  rq_init_comm_if_connected(9, "1")
  rq_init_comm_if_connected(2, "2")
  rq_init_comm_if_connected(3, "3")
  rq_init_comm_if_connected(4, "4")
  rq_print_connected_grippers()
  rq_gripper_communication_thread = run rq_gripper_communication()
  set_closed_norm(97.6470588235294, 1)
  set_open_norm(1.1764705882352942, 1)
  set_closed_mm(0.0, 1)
  set_open_mm(53.0, 1)
  set_closed_norm(100.0, 2)
  set_open_norm(0.0, 2)
  set_closed_mm(0.0, 2)
  set_open_mm(50.0, 2)
  set_closed_norm(100.0, 3)
  set_open_norm(0.0, 3)
  set_closed_mm(0.0, 3)
  set_open_mm(50.0, 3)
  set_closed_norm(100.0, 4)
  set_open_norm(0.0, 4)
  set_closed_mm(0.0, 4)
  set_open_mm(50.0, 4)
  rq_current_limit_enabled = False
  while(not rq_gripper_communication_thread_started):
      sync()
  end
  # end: URCap Installation Node
  global AMR_Position=struct(position_identifier=0, x1=0, x2=0, y1=0, y2=0, theta1=0, theta2=0)
  global CAM_Pose=p[0,0,0,0,0,0]
  global CAM_Relation=""
  global CMD_Abort=  False
  global CMD_Clear=  False
  global CMD_Reset=  False
  global CMD_Start=  False
  global CMD_Suspend=  False
  global CMD_Unhold=  False
  global CMD_Unsuspend=  False
  global CNT_Rack_Output=0
  global FNC_Freedrive=  False
  global PRC_TubCounter=0
  global PRC_TubNumber=0
  global STP=0
  global TMR_Barcode=0
  global TMR_Barcode_is_counting=False
  thread Timer_Thread():
    while (True):
      if (TMR_Barcode_is_counting):
        TMR_Barcode = TMR_Barcode + get_steptime()
      end
      sync()
    end
  end
  run Timer_Thread()
  def Sub_Vision_V18():
    $ 698 "Sub_Vision_V18" "noBreak"
    $ 699 "PreSettings"
    $ 700 "CAM_LM_Detected≔ False "
    global CAM_LM_Detected=  False
    $ 701 "CAM_Captures≔0"
    global CAM_Captures=0
    $ 702 "CAM_Pose≔p[0,0,0,0,0,0]"
    global CAM_Pose=p[0,0,0,0,0,0]
    $ 703 "CAM_LM_Refinmnt≔ False "
    global CAM_LM_Refinmnt=  False
    $ 704 "CAM_LM_Refined≔ False "
    global CAM_LM_Refined=  False
    $ 705 "CAM_LM_Deviatn≔p[0,0,0,0,0,0]"
    global CAM_LM_Deviatn=p[0,0,0,0,0,0]
    $ 706 "CAM_LM_ID≔0"
    global CAM_LM_ID=0
    $ 707 "CAM_Done≔ False "
    global CAM_Done=  False
    $ 708 "CAM_CNT_Obj≔0"
    global CAM_CNT_Obj=0
    $ 709 "CAM_Result = []"
    CAM_Result = []
    $ 710 "OBJ_Detected≔ False "
    global OBJ_Detected=  False
    $ 711 "FRM_Reference≔p[0,0,0,0,0,0]"
    global FRM_Reference=p[0,0,0,0,0,0]
    $ 712 "'=========='"
    # '=========='
    $ 713 "Switch Action"
    switch_1 = Action
    $ 714 "Case 13"
    if (13 == switch_1):
    elif (15 == switch_1):
      $ 832 "Case 15"
    elif (131 == switch_1):
      $ 878 "Case 131"
      $ 879 "Read (SensoPart)"
      $ 880 "Action_Info≔'search for landmark'"
      global Action_Info="search for landmark"
      $ 881 "CAM_LM≔CAM_LMs[ITM_ID-1]"
      global CAM_LM=CAM_LMs[ITM_ID-1]
      $ 882 "CAM_Relation≔CAM_LM.capture_relation"
      global CAM_Relation=CAM_LM.capture_relation
      $ 883 "go to capture pose"
      $ 886 "If ITM_ID≟1 and JIG≟7"
      if (ITM_ID == 1  and  JIG == 7):
        $ 887 "PSE_T≔uLM_Cap_SSRack"
        global PSE_T=uLM_Cap_SSRack
      else:
        $ 888 "ElseIf ITM_ID≟5 and JIG≟7"
        if (ITM_ID == 5  and  JIG == 7):
          $ 889 "PSE_T≔FRM_Cap_SSRack"
          global PSE_T=FRM_Cap_SSRack
        end
      end
      $ 890 "do_transition(PSE_T, keep_rxry=False)"
      do_transition(PSE_T, keep_rxry=False)
      $ 891 "Set"
      set_tcp(p[0.0,0.0,0.161,3.1415,0.0,0.0])
      $ 892 "MoveJ"
      $ 893 "PSE_T" "breakAfter"
      movej(PSE_T, a=1.3962634015954636, v=1.7453292519943295)
      $ 894 "CAM_Pose≔get_actual_tcp_pose()"
      global CAM_Pose= get_actual_tcp_pose ()
      $ 895 "Loop  not CAM_Done and  not ERROR.FLAG and  not CMD_Stop"
      while (  not  CAM_Done  and    not  ERROR.FLAG  and    not  CMD_Stop):
        $ 896 "adjust capture pose"
        $ 897 "If CAM_LM_Detected and CAM_LM_Refinmnt"
        if (CAM_LM_Detected  and  CAM_LM_Refinmnt):
          $ 898 "PSE_T≔p[0,0,0.300,0,0,0]"
          global PSE_T=p[0,0,0.300,0,0,0]
          $ 899 "CAM_Pose≔PSE_T"
          global CAM_Pose=PSE_T
          $ 900 "If  not is_reachable(FRM_Reference,[PSE_T])"
          if (  not  is_reachable(FRM_Reference,[PSE_T])):
            $ 901 "Error"
            $ 902 "set_error(ERROR_POSE_NOT_REACHABLE)"
            set_error(ERROR_POSE_NOT_REACHABLE)
          end
          $ 903 "If  not ERROR.FLAG"
          if (  not  ERROR.FLAG):
            $ 904 "MoveJ"
            $ 905 "PSE_T" "breakAfter"
            set_tcp(p[0.0,0.0,0.161,0.0,0.0,0.0])
            movej(pose_trans(FRM_Reference, PSE_T), a=0.8726646259971648, v=1.3962634015954636)
            $ 906 "CAM_LM_Refined≔ True "
            global CAM_LM_Refined=  True
          end
        else:
          $ 907 "ElseIf  not CAM_LM_Detected and CAM_Captures>0"
          if (  not  CAM_LM_Detected  and  CAM_Captures>0):
            $ 908 "MoveL"
            $ 909 "If FRM_Reference≟p[0,0,0,0,0,0]"
            if (FRM_Reference == p[0,0,0,0,0,0]):
              $ 910 "PSE_T≔get_random_pose(pose_ref=CAM_Pose, mode='cubic', range_max=[0.150,0.150,0.015])"
              global PSE_T=get_random_pose(pose_ref=CAM_Pose, mode="cubic", range_max=[0.150,0.150,0.015])
            else:
              $ 915 "Else" "noBreak"
              $ 916 "PSE_T≔get_random_pose(pose_ref=CAM_Pose, mode='rotation', range_max=[10,10,0])"
              global PSE_T=get_random_pose(pose_ref=CAM_Pose, mode="rotation", range_max=[10,10,0])
              $ 917 "CAM_LM_Refined≔ True "
              global CAM_LM_Refined=  True
            end
            $ 918 "If get_inverse_kin_has_solution(pose_trans(FRM_Reference, PSE_T))"
            if (get_inverse_kin_has_solution( pose_trans (FRM_Reference, PSE_T))):
              $ 919 "Comment"
              # Comment
              $ 920 "PSE_T" "breakAfter"
              set_tcp(p[0.0,0.0,0.161,3.1415,0.0,0.0])
              movel(pose_trans(FRM_Reference, PSE_T), a=0.03, v=0.05)
            else:
              $ 921 "Else" "noBreak"
              $ 922 "'If random pose is out of reach, set the initial cam pose'"
              # 'If random pose is out of reach, set the initial cam pose'
              $ 923 "PSE_T≔CAM_Pose"
              global PSE_T=CAM_Pose
            end
          end
        end
        $ 924 "Wait: 2.0"
        sleep(2.0)
        $ 925 "trigger"
        # begin: URCap Program Node
        #   Source: SensoPart VISOR Robotic, 2.0.0, SensoPart Industriesensorik GmbH
        #   Type: VISOR Trigger
        $ 926 "# 1 VISOR Trigger"
        visor_trigger(1, 6000, "arm")
        # end: URCap Program Node
        $ 930 "TM_3D_Found≔visor_partsFound(1)"
        global TM_3D_Found= visor_partsFound (1)
        $ 931 "If TM_3D_Found>0"
        if (TM_3D_Found>0):
          $ 932 "CAM_LM_Detected≔ True "
          global CAM_LM_Detected=  True
          $ 933 "CAM_Captures≔0"
          global CAM_Captures=0
        else:
          $ 934 "Else" "noBreak"
          $ 935 "CAM_LM_Detected≔ False "
          global CAM_LM_Detected=  False
          $ 936 "CAM_Captures≔CAM_Captures+1"
          global CAM_Captures=CAM_Captures+1
        end
        $ 941 "result"
        $ 942 "If CAM_LM_Detected"
        if (CAM_LM_Detected):
          $ 943 "If (CAM_LM_Refinmnt and CAM_LM_Refined) or  not CAM_LM_Refinmnt"
          if ((CAM_LM_Refinmnt  and  CAM_LM_Refined)  or    not  CAM_LM_Refinmnt):
            $ 1001 "If ITM_ID≟1 and JIG≟7"
            if (ITM_ID == 1  and  JIG == 7):
              $ 1002 "CAM_LM_SSRack≔visor_getPose3d(1, 0)"
              global CAM_LM_SSRack= visor_getPose3d (1, 0)
            else:
              $ 1003 "ElseIf ITM_ID≟5 and JIG≟7"
              if (ITM_ID == 5  and  JIG == 7):
                $ 1004 "CAM_LM_SSRack≔visor_getPose3d(1, 0)"
                global CAM_LM_SSRack= visor_getPose3d (1, 0)
              end
            end
            $ 1005 "CAM_Done≔ True "
            global CAM_Done=  True
          end
        else:
          $ 1006 "ElseIf  not CAM_LM_Detected and CAM_Captures<CAM_PRM_Retries"
          if (  not  CAM_LM_Detected  and  CAM_Captures<CAM_PRM_Retries):
            $ 1007 "CAM_LM_Refined≔ False "
            global CAM_LM_Refined=  False
          else:
            $ 1008 "ElseIf CAM_Captures≥CAM_PRM_Retries"
            if (CAM_Captures >= CAM_PRM_Retries):
              $ 1009 "CAM_Done≔ True "
              global CAM_Done=  True
              $ 1010 "Error"
              $ 1011 "set_error(ERROR_NO_LANDMARK)"
              set_error(ERROR_NO_LANDMARK)
            end
          end
        end
      end
    elif (151 == switch_1):
      $ 1012 "Case 151"
      $ 1013 "Detect (SensoPart)"
      $ 1014 "go to capture pose"
      $ 1015 "FRM_Reference≔FRM_Cap_SSRack"
      global FRM_Reference=FRM_Cap_SSRack
      $ 1016 "PSE_T≔p[0,0,-0.00,0,0,0]"
      global PSE_T=p[0,0,-0.00,0,0,0]
      $ 1017 "do_transition(pose_trans(FRM_Reference, PSE_T), keep_rxry=False)"
      do_transition( pose_trans (FRM_Reference, PSE_T), keep_rxry=False)
      $ 1018 "JNT_Q≔get_actual_joint_positions()"
      global JNT_Q= get_actual_joint_positions ()
      $ 1019 "JNT_Q≔[JNT_Q[0], JNT_Q[1], JNT_Q[2], JNT_Q[3], JNT_Q[4], 0]"
      global JNT_Q=[JNT_Q[0], JNT_Q[1], JNT_Q[2], JNT_Q[3], JNT_Q[4], 0]
      $ 1020 "Set"
      set_tcp(p[0.0,0.0,0.161,3.1415,0.0,0.0])
      $ 1021 "movej(get_inverse_kin(pose_trans(FRM_Reference, PSE_T), qnear=JNT_Q))"
      movej(get_inverse_kin( pose_trans (FRM_Reference, PSE_T), qnear=JNT_Q))
      $ 1022 "CAM_Pose≔pose_trans(pose_inv(FRM_Reference), get_actual_tcp_pose())"
      global CAM_Pose= pose_trans ( pose_inv (FRM_Reference),  get_actual_tcp_pose ())
      $ 1023 "Loop  not CAM_Done and  not ERROR.FLAG and  not CMD_Stop"
      while (  not  CAM_Done  and    not  ERROR.FLAG  and    not  CMD_Stop):
        $ 1024 "If  not OBJ_Detected and CAM_Captures>0"
        if (  not  OBJ_Detected  and  CAM_Captures>0):
          $ 1025 "MoveL"
          $ 1026 "If FRM_Reference≟p[0,0,0,0,0,0]"
          if (FRM_Reference == p[0,0,0,0,0,0]):
            $ 1028 "PSE_T≔get_random_pose(pose_ref=CAM_Pose, mode='rotation', range_max=[15,15,0])"
            global PSE_T=get_random_pose(pose_ref=CAM_Pose, mode="rotation", range_max=[15,15,0])
          else:
            $ 1029 "Else" "noBreak"
            $ 1030 "PSE_T≔get_random_pose(pose_ref=CAM_Pose, mode='rotation', range_max=[10,10,0])"
            global PSE_T=get_random_pose(pose_ref=CAM_Pose, mode="rotation", range_max=[10,10,0])
          end
          $ 1031 "If get_inverse_kin_has_solution(pose_trans(FRM_Reference, PSE_T))"
          if (get_inverse_kin_has_solution( pose_trans (FRM_Reference, PSE_T))):
            $ 1032 "PSE_T" "breakAfter"
            set_tcp(p[0.0,0.0,0.161,3.1415,0.0,0.0])
            movel(pose_trans(FRM_Reference, PSE_T), a=0.03, v=0.05)
          else:
            $ 1033 "Else" "noBreak"
            $ 1034 "'If random pose is out of reach, set the initial cam pose'"
            # 'If random pose is out of reach, set the initial cam pose'
            $ 1035 "PSE_T≔CAM_Pose"
            global PSE_T=CAM_Pose
            $ 1036 "PSE_T" "breakAfter"
            set_tcp(p[0.0,0.0,0.161,3.1415,0.0,0.0])
            movel(pose_trans(FRM_Reference, PSE_T), a=0.03, v=0.05)
          end
        end
        $ 1037 "Wait: 0.5"
        sleep(0.5)
        $ 1038 "Set"
        set_tcp(p[0.0,0.0,0.161,3.1415,0.0,0.0])
        # begin: URCap Program Node
        #   Source: SensoPart VISOR Robotic, 2.0.0, SensoPart Industriesensorik GmbH
        #   Type: VISOR Trigger
        $ 1039 "# 1 VISOR Trigger"
        visor_changeJob(1, "Object Detection Single", 6000)
        visor_trigger(1, 6000, "arm")
        # end: URCap Program Node
        $ 1040 "If visor_isResponseOk(1)"
        if ( visor_isResponseOk (1)):
          $ 1041 "CAM_CNT_Obj≔visor_partsFound(1)"
          global CAM_CNT_Obj= visor_partsFound (1)
          $ 1042 "CAM_OBJ_Pose≔visor_getPose3d(1, 0)"
          global CAM_OBJ_Pose= visor_getPose3d (1, 0)
          $ 1043 "If CAM_CNT_Obj>0"
          if (CAM_CNT_Obj>0):
            $ 1044 "CAM_OBJ_Color≔visor_getAdditionalData(1, 0)"
            global CAM_OBJ_Color= visor_getAdditionalData (1, 0)
            $ 1045 "CAM_DetectScore≔to_num(visor_getAdditionalData(1, 1))/1000"
            global CAM_DetectScore=to_num( visor_getAdditionalData (1, 1))/1000
            $ 1046 "OBJ_Detected≔ True "
            global OBJ_Detected=  True
          end
        else:
          $ 1047 "Else" "noBreak"
          $ 1048 "CAM_Captures≔CAM_Captures+1"
          global CAM_Captures=CAM_Captures+1
        end
        $ 1049 "If OBJ_Detected"
        if (OBJ_Detected):
          $ 1050 "Get object data"
          $ 1051 "PRC_CntDetect≔0"
          global PRC_CntDetect=0
          $ 1052 "Loop PRC_CntDetect<CAM_CNT_Obj"
          while (PRC_CntDetect<CAM_CNT_Obj):
            $ 1053 "get object and jig number"
            $ 1054 "If ITM_ID≟1 and JIG≟7"
            if (ITM_ID == 1  and  JIG == 7):
              $ 1055 "FRM_Reference≔FRM_Cap_SSRack"
              global FRM_Reference=FRM_Cap_SSRack
            else:
              $ 1056 "ElseIf ITM_ID≟5 and JIG≟7"
              if (ITM_ID == 5  and  JIG == 7):
                $ 1057 "FRM_Reference≔uLM_Cap_SSRack"
                global FRM_Reference=uLM_Cap_SSRack
              end
            end
            $ 1060 "PSE_T≔pose_trans(pose_inv(FRM_Reference), CAM_OBJ_Pose)"
            global PSE_T= pose_trans ( pose_inv (FRM_Reference), CAM_OBJ_Pose)
            $ 1061 "CAM_Result.append(get_pattern_counter(PSE_T, 'X', pattern=[10, 5], patternsize=[0.181, 0.081]))"
            CAM_Result.append(get_pattern_counter(PSE_T, "X", pattern=[10, 5], patternsize=[0.181, 0.081]))
            $ 1062 "PRC_CntDetect≔PRC_CntDetect+1"
            global PRC_CntDetect=PRC_CntDetect+1
          end
          $ 1063 "CAM_Done≔ True "
          global CAM_Done=  True
        else:
          $ 1064 "ElseIf CAM_Captures≥CAM_PRM_Retries"
          if (CAM_Captures >= CAM_PRM_Retries):
            $ 1065 "CAM_Done≔ True "
            global CAM_Done=  True
          else:
            $ 1066 "Else" "noBreak"
            $ 1067 "CAM_Captures≔CAM_Captures+1"
            global CAM_Captures=CAM_Captures+1
          end
        end
      end
    end
    $ 1068 "'=========='"
    # '=========='
    $ 1069 "PostSettings"
    $ 1070 "FRM_Reference≔p[0,0,0,0,0,0]"
    global FRM_Reference=p[0,0,0,0,0,0]
    $ 1071 "Set"
    set_tcp(p[0.0,0.0,0.161,3.1415,0.0,0.0])
    $ 1072 "CAM_Pose≔p[0,0,0,0,0,0]"
    global CAM_Pose=p[0,0,0,0,0,0]
    $ 1073 "Action≔0"
    global Action=0
    $ 1074 "Action_Info≔''"
    global Action_Info=""
  end
  def Sub_AMR_MiR_V3():
    $ 1075 "Sub_AMR_MiR_V3" "noBreak"
    $ 1076 "PreSettings"
    $ 1077 "AMR_TargetList≔[1,2,3,4,5,21,22,23,24,31,32,33,34,35,36,37,38,41]"
    global AMR_TargetList=[1,2,3,4,5,21,22,23,24,31,32,33,34,35,36,37,38,41]
    $ 1078 "AMR_Done≔ False "
    global AMR_Done=  False
    $ 1079 "AMR_PosActual≔T2O_Current_Pos"
    global AMR_PosActual=modbus_get_signal_status("T2O_Current_Pos")
    $ 1080 "AMR_Attemps≔T2O_Nav_Attemps"
    global AMR_Attemps=modbus_get_signal_status("T2O_Nav_Attemps")
    $ 1081 "AMR_Battery≔MiR_Battery_Lvl"
    global AMR_Battery=modbus_get_signal_status("MiR_Battery_Lvl")
    $ 1082 "AMR_Charging≔(T2O_Charging≟1)"
    global AMR_Charging=(modbus_get_signal_status("T2O_Charging") == 1)
    $ 1083 "AMR_Position≔struct(position_identifier=T2O_Current_Pos, x1=MiR_Position_X1, x2=MiR_Position_X2, y1=MiR_Position_Y1, y2=MiR_Position_Y2, theta1=MiR_Theta_1, theta2=MiR_Theta_2) "
    global AMR_Position=struct(position_identifier=modbus_get_signal_status("T2O_Current_Pos"), x1=modbus_get_signal_status("MiR_Position_X1"), x2=modbus_get_signal_status("MiR_Position_X2"), y1=modbus_get_signal_status("MiR_Position_Y1"), y2=modbus_get_signal_status("MiR_Position_Y2"), theta1=modbus_get_signal_status("MiR_Theta_1"), theta2=modbus_get_signal_status("MiR_Theta_2"))
    $ 1084 "If MiR_Mode≠7"
    if (modbus_get_signal_status("MiR_Mode") != 7):
      $ 1085 "Error"
      $ 1086 "set_error(ERROR_AMR_WRONG_MODE)"
      set_error(ERROR_AMR_WRONG_MODE)
      $ 1087 "AMR_Done≔ True "
      global AMR_Done=  True
    end
    $ 1088 "'=========='"
    # '=========='
    $ 1089 "Switch STATE"
    switch_1 = STATE
    $ 1090 "Case 1"
    if (1 == switch_1):
      $ 1091 "stopping"
      $ 1092 "If T2O_Done≟1 and O2T_Acknowledge≟0"
      if (modbus_get_signal_status("T2O_Done") == 1  and  modbus_get_signal_status("O2T_Acknowledge") == 0):
        $ 1093 "Set O2T_Acknowledge=1"
        modbus_set_output_register("O2T_Acknowledge", 1)
      end
      $ 1094 "Set MiR_CMD_Stop=On"
      modbus_set_output_signal("MiR_CMD_Stop", True)
      $ 1095 "AMR_Position.position_identifier = 0"
      AMR_Position.position_identifier = 0
      $ 1096 "AMR_Done≔ True "
      global AMR_Done=  True
    elif (2 == switch_1):
      $ 1097 "Case 2"
      $ 1098 "stopped"
      $ 1099 "If MiR_State≠3 and MiR_State≠5"
      if (modbus_get_signal_status("MiR_State") != 3  and  modbus_get_signal_status("MiR_State") != 5):
        $ 1100 "Set MiR_CMD_Stop=Off"
        modbus_set_output_signal("MiR_CMD_Stop", False)
      end
    elif (3 == switch_1):
      $ 1101 "Case 3"
      $ 1102 "resetting"
      $ 1103 "Set O2T_Mis_Main=Off"
      modbus_set_output_signal("O2T_Mis_Main", False)
      $ 1104 "Set O2T_Mis_Charge=Off"
      modbus_set_output_signal("O2T_Mis_Charge", False)
      $ 1105 "If MiR_Mis_Queue>0"
      if (modbus_get_signal_status("MiR_Mis_Queue")>0):
        $ 1106 "Set MiR_CMD_Clear_Q=On"
        modbus_set_output_signal("MiR_CMD_Clear_Q", True)
        $ 1107 "Wait MiR_Mis_Queue≟0"
        while (not(modbus_get_signal_status("MiR_Mis_Queue") == 0)):
          sync()
        end
        $ 1108 "Set MiR_CMD_Clear_Q=Off"
        modbus_set_output_signal("MiR_CMD_Clear_Q", False)
      end
      $ 1109 "If MiR_Error_ID≠0"
      if (modbus_get_signal_status("MiR_Error_ID") != 0):
        $ 1110 "Set MiR_CMD_Clear_E=On"
        modbus_set_output_signal("MiR_CMD_Clear_E", True)
        $ 1111 "Wait MiR_Error_ID≟0"
        while (not(modbus_get_signal_status("MiR_Error_ID") == 0)):
          sync()
        end
        $ 1112 "Set MiR_CMD_Clear_E=Off"
        modbus_set_output_signal("MiR_CMD_Clear_E", False)
      end
      $ 1113 "Set O2T_Action=0"
      modbus_set_output_register("O2T_Action", 0)
      $ 1114 "Set O2T_Acknowledge=0"
      modbus_set_output_register("O2T_Acknowledge", 0)
      $ 1115 "Set O2T_Target_Pos=0"
      modbus_set_output_register("O2T_Target_Pos", 0)
      $ 1116 "Set O2T_Footprint=0"
      modbus_set_output_register("O2T_Footprint", 0)
      $ 1117 "Set O2T_ProtectOff=0"
      modbus_set_output_register("O2T_ProtectOff", 0)
      $ 1118 "Set O2T_Dock=0"
      modbus_set_output_register("O2T_Dock", 0)
      $ 1119 "AMR_Attemps≔0"
      global AMR_Attemps=0
      $ 1120 "AMR_PosTarget≔0"
      global AMR_PosTarget=0
      $ 1121 "AMR_Step≔0"
      global AMR_Step=0
      $ 1122 "AMR_AtTarget≔ False "
      global AMR_AtTarget=  False
      $ 1123 "If MiR_State≟4 or MiR_State≟3 or MiR_State≟10"
      if (modbus_get_signal_status("MiR_State") == 4  or  modbus_get_signal_status("MiR_State") == 3  or  modbus_get_signal_status("MiR_State") == 10):
        $ 1124 "AMR_Done≔ True "
        global AMR_Done=  True
      end
    elif (5 == switch_1):
      $ 1125 "Case 5"
      $ 1126 "starting"
      $ 1127 "If MiR_State≟4"
      if (modbus_get_signal_status("MiR_State") == 4):
        $ 1128 "Set MiR_CMD_Start=On"
        modbus_set_output_signal("MiR_CMD_Start", True)
        $ 1129 "Wait MiR_State≠4"
        while (not(modbus_get_signal_status("MiR_State") != 4)):
          sync()
        end
        $ 1130 "Set MiR_CMD_Start=Off"
        modbus_set_output_signal("MiR_CMD_Start", False)
        $ 1131 "AMR_Done≔ True "
        global AMR_Done=  True
      else:
        $ 1132 "ElseIf MiR_State≟10"
        if (modbus_get_signal_status("MiR_State") == 10):
          $ 1133 "'MiR in protective stop. Wait'"
          # 'MiR in protective stop. Wait'
          $ 1134 "AMR_Done≔ True "
          global AMR_Done=  True
        else:
          $ 1135 "ElseIf MiR_State≟3"
          if (modbus_get_signal_status("MiR_State") == 3):
            $ 1136 "AMR_Done≔ True "
            global AMR_Done=  True
          end
        end
      end
    elif (6 == switch_1):
      $ 1137 "Case 6"
      $ 1138 "execute"
      $ 1139 "AMR_AtTarget≔(AMR_PosActual≟AMR_PosTarget)"
      global AMR_AtTarget=(AMR_PosActual == AMR_PosTarget)
      $ 1140 "Switch AMR_Step"
      switch_2 = AMR_Step
      $ 1141 "Case 0"
      if (0 == switch_2):
        $ 1142 "If  not AMR_AtTarget"
        if (  not  AMR_AtTarget):
          $ 1143 "AMR_Step≔1"
          global AMR_Step=1
        else:
          $ 1144 "Else" "noBreak"
          $ 1145 "AMR_Done≔ True "
          global AMR_Done=  True
        end
      elif (1 == switch_2):
        $ 1146 "Case 1"
        $ 1147 "general Settings"
        $ 1148 "Set O2T_Acknowledge=0"
        modbus_set_output_register("O2T_Acknowledge", 0)
        $ 1149 "check for error"
        $ 1150 "If OBJ_Picked and MiR_State≟10"
        if (OBJ_Picked  and  modbus_get_signal_status("MiR_State") == 10):
          $ 1151 "Error"
          $ 1152 "set_error(ERROR_ROBOT_ARM_NOT_IN_HOME_POSE)"
          set_error(ERROR_ROBOT_ARM_NOT_IN_HOME_POSE)
          $ 1153 "Action≔0"
          global Action=0
        else:
          $ 1154 "ElseIf  not found_in_list(AMR_PosTarget, AMR_TargetList)"
          if (  not  found_in_list(AMR_PosTarget, AMR_TargetList)):
            $ 1155 "Error"
            $ 1156 "set_error(ERROR_UNKNOWN_POSE)"
            set_error(ERROR_UNKNOWN_POSE)
            $ 1157 "Action≔0"
            global Action=0
          end
        end
        $ 1158 "If MiR_State≟3"
        if (modbus_get_signal_status("MiR_State") == 3):
          $ 1159 "Set MiR_CMD_Start=Off"
          modbus_set_output_signal("MiR_CMD_Start", False)
          $ 1160 "Switch Action"
          switch_3 = Action
          $ 1161 "Case 51"
          if (51 == switch_3):
            $ 1162 "Charge"
            $ 1163 "'trigger the charging mission'"
            # 'trigger the charging mission'
            $ 1164 "'target pos is predefined'"
            # 'target pos is predefined'
            $ 1165 "Set O2T_Footprint=0"
            modbus_set_output_register("O2T_Footprint", 0)
            $ 1166 "Set O2T_Action=1"
            modbus_set_output_register("O2T_Action", 1)
            $ 1167 "If MiR_Mis_Queue≟0"
            if (modbus_get_signal_status("MiR_Mis_Queue") == 0):
              $ 1168 "Set O2T_Mis_Charge=On"
              modbus_set_output_signal("O2T_Mis_Charge", True)
              $ 1169 "Wait MiR_Mis_Queue≥1"
              while (not(modbus_get_signal_status("MiR_Mis_Queue") >= 1)):
                sync()
              end
              $ 1170 "Set O2T_Mis_Charge=Off"
              modbus_set_output_signal("O2T_Mis_Charge", False)
            end
          elif (52 == switch_3):
            $ 1171 "Case 52"
            $ 1172 "Navigate"
            $ 1173 "'trigger the standard missoin'"
            # 'trigger the standard missoin'
            $ 1174 "Set O2T_Footprint=AMR_FootprintID"
            modbus_set_output_register("O2T_Footprint", AMR_FootprintID)
            $ 1175 "Set O2T_Target_Pos=AMR_PosTarget"
            modbus_set_output_register("O2T_Target_Pos", AMR_PosTarget)
            $ 1176 "Set O2T_Action=2"
            modbus_set_output_register("O2T_Action", 2)
            $ 1177 "If MiR_Mis_Queue≟0"
            if (modbus_get_signal_status("MiR_Mis_Queue") == 0):
              $ 1178 "Set O2T_Mis_Main=On"
              modbus_set_output_signal("O2T_Mis_Main", True)
              $ 1179 "Wait MiR_Mis_Queue≥1"
              while (not(modbus_get_signal_status("MiR_Mis_Queue") >= 1)):
                sync()
              end
              $ 1180 "Set O2T_Mis_Main=Off"
              modbus_set_output_signal("O2T_Mis_Main", False)
            end
          end
        else:
          $ 1181 "ElseIf MiR_State≟4"
          if (modbus_get_signal_status("MiR_State") == 4):
            $ 1182 "Set MiR_CMD_Start=On"
            modbus_set_output_signal("MiR_CMD_Start", True)
          else:
            $ 1183 "ElseIf MiR_State≟5"
            if (modbus_get_signal_status("MiR_State") == 5):
              $ 1184 "AMR_Step≔2"
              global AMR_Step=2
            else:
              $ 1185 "ElseIf MiR_State≟10"
              if (modbus_get_signal_status("MiR_State") == 10):
                $ 1186 "'AMR still in safeguard stop'"
                # 'AMR still in safeguard stop'
              end
            end
          end
        end
      elif (2 == switch_2):
        $ 1187 "Case 2"
        $ 1188 "acknowledge handshake"
        $ 1189 "If T2O_Done≟1 and O2T_Acknowledge≟0"
        if (modbus_get_signal_status("T2O_Done") == 1  and  modbus_get_signal_status("O2T_Acknowledge") == 0):
          $ 1190 "Set O2T_Acknowledge=1"
          modbus_set_output_register("O2T_Acknowledge", 1)
        else:
          $ 1191 "ElseIf T2O_Done≟0 and O2T_Acknowledge≟1"
          if (modbus_get_signal_status("T2O_Done") == 0  and  modbus_get_signal_status("O2T_Acknowledge") == 1):
            $ 1192 "Set O2T_Acknowledge=0"
            modbus_set_output_register("O2T_Acknowledge", 0)
            $ 1193 "AMR_AtTarget≔(AMR_PosActual≟AMR_PosTarget)"
            global AMR_AtTarget=(AMR_PosActual == AMR_PosTarget)
            $ 1194 "AMR_Done≔ True "
            global AMR_Done=  True
          end
        end
      end
      $ 1195 "translate errors"
      $ 1196 "If AMR_Done"
      if (AMR_Done):
        $ 1197 "Switch T2O_Error_ID"
        switch_2 = modbus_get_signal_status("T2O_Error_ID")
        $ 1198 "Case 2003"
        if (2003 == switch_2):
          $ 1199 "error"
          $ 1200 "set_error(ERROR_NOT_DOCKED)"
          set_error(ERROR_NOT_DOCKED)
        elif (2007 == switch_2):
          $ 1201 "Case 2007"
          $ 1202 "error"
          $ 1203 "set_error(ERROR_NOT_REACHABLE_TARGET)"
          set_error(ERROR_NOT_REACHABLE_TARGET)
        elif (2008 == switch_2):
          $ 1204 "Case 2008"
          $ 1205 "error"
          $ 1206 "set_error(ERROR_CHARGING_NOT_STARTED)"
          set_error(ERROR_CHARGING_NOT_STARTED)
        end
      end
    elif (7 == switch_1):
      $ 1207 "Case 7"
      $ 1208 "completing"
      $ 1209 "If MiR_Mis_Queue>0"
      if (modbus_get_signal_status("MiR_Mis_Queue")>0):
        $ 1210 "Set MiR_CMD_Abort=On"
        modbus_set_output_signal("MiR_CMD_Abort", True)
        $ 1211 "Wait MiR_Mis_Queue≟0"
        while (not(modbus_get_signal_status("MiR_Mis_Queue") == 0)):
          sync()
        end
        $ 1212 "Set MiR_CMD_Abort=Off"
        modbus_set_output_signal("MiR_CMD_Abort", False)
      end
      $ 1213 "If MiR_State≟3 or MiR_State≟10"
      if (modbus_get_signal_status("MiR_State") == 3  or  modbus_get_signal_status("MiR_State") == 10):
        $ 1214 "AMR_Done≔ True "
        global AMR_Done=  True
      end
    elif (9 == switch_1):
      $ 1215 "Case 9"
      $ 1216 "holding"
      $ 1217 "Set MiR_CMD_Abort=On"
      modbus_set_output_signal("MiR_CMD_Abort", True)
      $ 1218 "If MiR_State≟3 or MiR_State≟10"
      if (modbus_get_signal_status("MiR_State") == 3  or  modbus_get_signal_status("MiR_State") == 10):
        $ 1219 "Set MiR_CMD_Abort=Off"
        modbus_set_output_signal("MiR_CMD_Abort", False)
        $ 1220 "AMR_Done≔ True "
        global AMR_Done=  True
      end
    elif (11 == switch_1):
      $ 1221 "Case 11"
      $ 1222 "unholding"
      $ 1223 "Set MiR_CMD_Start=On"
      modbus_set_output_signal("MiR_CMD_Start", True)
      $ 1224 "If MiR_State≠4"
      if (modbus_get_signal_status("MiR_State") != 4):
        $ 1225 "Set MiR_CMD_Start=Off"
        modbus_set_output_signal("MiR_CMD_Start", False)
        $ 1226 "AMR_Step≔0"
        global AMR_Step=0
        $ 1227 "AMR_Done≔ True "
        global AMR_Done=  True
      end
    elif (12 == switch_1):
      $ 1228 "Case 12"
      $ 1229 "suspending"
      $ 1230 "'none'"
      # 'none'
    elif (14 == switch_1):
      $ 1231 "Case 14"
      $ 1232 "unsuspending"
      $ 1233 "'none'"
      # 'none'
    elif (15 == switch_1):
      $ 1234 "Case 15"
      $ 1235 "aborting"
      $ 1236 "Set MiR_CMD_Abort=On"
      modbus_set_output_signal("MiR_CMD_Abort", True)
      $ 1237 "Wait MiR_State≟3"
      while (not(modbus_get_signal_status("MiR_State") == 3)):
        sync()
      end
      $ 1238 "Set MiR_CMD_Abort=Off"
      modbus_set_output_signal("MiR_CMD_Abort", False)
    elif (17 == switch_1):
      $ 1239 "Case 17"
      $ 1240 "clearing"
      $ 1241 "If MiR_Error_ID≠0"
      if (modbus_get_signal_status("MiR_Error_ID") != 0):
        $ 1242 "Set MiR_CMD_Clear_E=On"
        modbus_set_output_signal("MiR_CMD_Clear_E", True)
        $ 1243 "Wait MiR_Error_ID≟0"
        while (not(modbus_get_signal_status("MiR_Error_ID") == 0)):
          sync()
        end
        $ 1244 "Set MiR_CMD_Clear_E=Off"
        modbus_set_output_signal("MiR_CMD_Clear_E", False)
      end
      $ 1245 "If MiR_Error_ID≟0"
      if (modbus_get_signal_status("MiR_Error_ID") == 0):
        $ 1246 "AMR_Done≔ True "
        global AMR_Done=  True
      end
    end
    $ 1247 "'=========='"
    # '=========='
    $ 1248 "PostSettings"
    $ 1249 "AMR_Position≔struct(position_identifier=T2O_Current_Pos, x1=MiR_Position_X1, x2=MiR_Position_X2, y1=MiR_Position_Y1, y2=MiR_Position_Y2, theta1=MiR_Theta_1, theta2=MiR_Theta_2) "
    global AMR_Position=struct(position_identifier=modbus_get_signal_status("T2O_Current_Pos"), x1=modbus_get_signal_status("MiR_Position_X1"), x2=modbus_get_signal_status("MiR_Position_X2"), y1=modbus_get_signal_status("MiR_Position_Y1"), y2=modbus_get_signal_status("MiR_Position_Y2"), theta1=modbus_get_signal_status("MiR_Theta_1"), theta2=modbus_get_signal_status("MiR_Theta_2"))
  end
  def Sub_Action_V4():
    $ 1250 "Sub_Action_V4" "noBreak"
    $ 1251 "PreSettings"
    $ 1252 "init poses"
    $ 1253 "PSE_A≔p[0,0,0,0,0,0]"
    global PSE_A=p[0,0,0,0,0,0]
    $ 1254 "PSE_A_H≔p[0,0,0,0,0,0]"
    global PSE_A_H=p[0,0,0,0,0,0]
    $ 1255 "PSE_T≔p[0,0,0,0,0,0]"
    global PSE_T=p[0,0,0,0,0,0]
    $ 1256 "PSE_T_H≔p[0,0,0,0,0,0]"
    global PSE_T_H=p[0,0,0,0,0,0]
    $ 1257 "PSE_G≔p[0,0,0,0,0,0]"
    global PSE_G=p[0,0,0,0,0,0]
    $ 1258 "PSE_G_H≔p[0,0,0,0,0,0]"
    global PSE_G_H=p[0,0,0,0,0,0]
    $ 1259 "PSE_R≔p[0,0,0,0,0,0]"
    global PSE_R=p[0,0,0,0,0,0]
    $ 1260 "PSE_R_H≔p[0,0,0,0,0,0]"
    global PSE_R_H=p[0,0,0,0,0,0]
    $ 1261 "JNT_Q≔[0,0,0,0,0,0]"
    global JNT_Q=[0,0,0,0,0,0]
    $ 1262 "JNT_S≔[0,0,0,0,0,0]"
    global JNT_S=[0,0,0,0,0,0]
    $ 1263 "Gripping parameters"
    $ 1264 "OBJ = find_object_by_type(OBJs, OBJ_Type)"
    OBJ = find_object_by_type(OBJs, OBJ_Type)
    $ 1265 "GRP_Open_Pos≔OBJ.dimension.diameter * 1000 + 6"
    global GRP_Open_Pos=OBJ.dimension.diameter * 1000 + 6
    $ 1266 "GRP_Offset≔OBJ.gripper_offset"
    global GRP_Offset=OBJ.gripper_offset
    $ 1267 "rq_set_force_norm(50)"
     rq_set_force_norm (50)
    $ 1268 "rq_set_speed_norm(50)"
     rq_set_speed_norm (50)
    $ 1269 "Switch ITM_ID"
    switch_1 = ITM_ID
    $ 1270 "Case 1"
    if (1 == switch_1):
      $ 1271 "uML"
      $ 1272 "JIG2 = find_object_by_type(JIGs, JIG)"
      JIG2 = find_object_by_type(JIGs, JIG)
      $ 1273 "JIG_Offset≔JIG2.jig_offset"
      global JIG_Offset=JIG2.jig_offset
      $ 1274 "Switch JIG"
      switch_2 = JIG
      $ 1275 "Case 1"
      if (1 == switch_2):
        $ 1276 "3FG"
        $ 1277 "define poses"
        $ 1278 "FRM_Reference≔ULM_3FG"
        global FRM_Reference=ULM_3FG
        $ 1279 "JNT_Q≔JNT_HOME"
        global JNT_Q=JNT_HOME
        $ 1280 "PSE_T≔pose_trans(GRP_Offset, JIG_Offset)"
        global PSE_T= pose_trans (GRP_Offset, JIG_Offset)
        $ 1281 "PSE_A≔pose_trans(PSE_T, p[0,0,0.100,0,0,0])"
        global PSE_A= pose_trans (PSE_T, p[0,0,0.100,0,0,0])
        $ 1282 "PSE_R≔pose_add(PSE_T, p[0,0,0.100,0,0,0])"
        global PSE_R= pose_add (PSE_T, p[0,0,0.100,0,0,0])
      elif (2 == switch_2):
        $ 1283 "Case 2"
        $ 1284 "Input"
        $ 1285 "'CHANGE THE REFERENCE TO THE FRAME TO MOVE IN'"
        # 'CHANGE THE REFERENCE TO THE FRAME TO MOVE IN'
        $ 1286 "define poses"
        $ 1287 "FRM_Reference≔ULM_Input"
        global FRM_Reference=ULM_Input
        $ 1288 "PSE_T≔pose_trans(pose_trans(get_pattern_pos_rectangle(OBJ_Nbr, 'X', [10,5], patternsize=[0.181,0.081]), GRP_Offset), JIG_Offset)"
        global PSE_T= pose_trans ( pose_trans (get_pattern_pos_rectangle(OBJ_Nbr, "X", [10,5], patternsize=[0.181,0.081]), GRP_Offset), JIG_Offset)
        $ 1289 "If Action≟1"
        if (Action == 1):
          $ 1290 "PSE_R≔pose_add(PSE_T, p[0,0,0.200,0,0,0])"
          global PSE_R= pose_add (PSE_T, p[0,0,0.200,0,0,0])
          $ 1291 "PSE_A≔pose_add(PSE_T, p[0,0,0.100,0,0,0])"
          global PSE_A= pose_add (PSE_T, p[0,0,0.100,0,0,0])
        else:
          $ 1292 "ElseIf Action≟2"
          if (Action == 2):
            $ 1293 "PSE_R≔pose_add(PSE_T, p[0,0,0.100,0,0,0])"
            global PSE_R= pose_add (PSE_T, p[0,0,0.100,0,0,0])
            $ 1294 "PSE_A≔pose_add(PSE_T, p[0,0,0.200,0,0,0])"
            global PSE_A= pose_add (PSE_T, p[0,0,0.200,0,0,0])
          end
        end
      elif (3 == switch_2):
        $ 1295 "Case 3"
        $ 1296 "Output"
        $ 1297 "'CHANGE THE REFERENCE TO THE FRAME TO MOVE IN'"
        # 'CHANGE THE REFERENCE TO THE FRAME TO MOVE IN'
        $ 1298 "define poses"
        $ 1299 "FRM_Reference≔ULM_Output"
        global FRM_Reference=ULM_Output
        $ 1300 "PSE_T≔pose_trans(pose_trans(get_pattern_pos_rectangle(OBJ_Nbr, 'X', [10,5], patternsize=[0.181,0.081]), GRP_Offset), JIG_Offset)"
        global PSE_T= pose_trans ( pose_trans (get_pattern_pos_rectangle(OBJ_Nbr, "X", [10,5], patternsize=[0.181,0.081]), GRP_Offset), JIG_Offset)
        $ 1302 "If Action≟1"
        if (Action == 1):
          $ 1303 "PSE_R≔pose_add(PSE_T, p[0,0,0.200,0,0,0])"
          global PSE_R= pose_add (PSE_T, p[0,0,0.200,0,0,0])
          $ 1304 "PSE_A≔pose_add(PSE_T, p[0,0,0.100,0,0,0])"
          global PSE_A= pose_add (PSE_T, p[0,0,0.100,0,0,0])
        else:
          $ 1305 "ElseIf Action≟2"
          if (Action == 2):
            $ 1306 "PSE_R≔pose_add(PSE_T, p[0,0,0.100,0,0,0])"
            global PSE_R= pose_add (PSE_T, p[0,0,0.100,0,0,0])
            $ 1307 "PSE_A≔pose_add(PSE_T, p[0,0,0.200,0,0,0])"
            global PSE_A= pose_add (PSE_T, p[0,0,0.200,0,0,0])
          end
        end
      elif (4 == switch_2):
        $ 1308 "Case 4"
        $ 1309 "jig centrifuge racks"
        $ 1310 "define poses"
        $ 1311 "FRM_Reference≔ULM_Cent_Racks"
        global FRM_Reference=ULM_Cent_Racks
        $ 1312 "PSE_T≔get_pattern_pos_rectangle(JIG_Slot, 'X', [4,1], patternsize=[0.291,0])"
        global PSE_T=get_pattern_pos_rectangle(JIG_Slot, "X", [4,1], patternsize=[0.291,0])
        $ 1313 "If OBJ_Nbr≠0"
        if (OBJ_Nbr != 0):
          $ 1314 "PSE_T≔pose_trans(pose_trans(PSE_T, get_pattern_pos_rectangle(OBJ_Nbr, 'X', [3,3], patternsize=[0.060,0.060])),p[-0.030, -0.030,0,0,0,3.927])"
          global PSE_T= pose_trans ( pose_trans (PSE_T, get_pattern_pos_rectangle(OBJ_Nbr, "X", [3,3], patternsize=[0.060,0.060])),p[-0.030, -0.030,0,0,0,3.927])
        end
        $ 1315 "PSE_T≔pose_trans(PSE_T, GRP_Offset)"
        global PSE_T= pose_trans (PSE_T, GRP_Offset)
        $ 1316 "If Action≟1"
        if (Action == 1):
          $ 1317 "PSE_R≔pose_add(PSE_T, p[0,0,0.200,0,0,0])"
          global PSE_R= pose_add (PSE_T, p[0,0,0.200,0,0,0])
          $ 1318 "PSE_A≔pose_add(PSE_T, p[0,0,0.100,0,0,0])"
          global PSE_A= pose_add (PSE_T, p[0,0,0.100,0,0,0])
        else:
          $ 1319 "ElseIf Action≟2"
          if (Action == 2):
            $ 1320 "PSE_R≔pose_add(PSE_T, p[0,0,0.100,0,0,0])"
            global PSE_R= pose_add (PSE_T, p[0,0,0.100,0,0,0])
            $ 1321 "PSE_A≔pose_add(PSE_T, p[0,0,0.200,0,0,0])"
            global PSE_A= pose_add (PSE_T, p[0,0,0.200,0,0,0])
          end
        end
      elif (6 == switch_2):
        $ 1322 "Case 6"
        $ 1323 "Caps bin"
        $ 1324 "define poses"
        $ 1325 "'Drop cap'"
        # 'Drop cap'
        $ 1326 "FRM_Reference=ULM_Cap_Bin"
        FRM_Reference=ULM_Cap_Bin
        $ 1327 "PSE_T≔pose_RPY2RotVec(p[0,0,0,0,0,0])"
        global PSE_T=pose_RPY2RotVec(p[0,0,0,0,0,0])
        $ 1328 "PSE_T_H≔pose_add(PSE_T, p[0,0,-0.011,0,0,0])"
        global PSE_T_H= pose_add (PSE_T, p[0,0,-0.011,0,0,0])
        $ 1329 "PSE_A≔pose_trans(PSE_T, p[0,0,0.1,0,0,0])"
        global PSE_A= pose_trans (PSE_T, p[0,0,0.1,0,0,0])
        $ 1330 "PSE_R_H≔pose_add(PSE_T, p[0,0,0.100,0,0,0])"
        global PSE_R_H= pose_add (PSE_T, p[0,0,0.100,0,0,0])
        $ 1331 "PSE_R≔pose_add(PSE_T, p[0,0,0.100,0,0,0])"
        global PSE_R= pose_add (PSE_T, p[0,0,0.100,0,0,0])
      elif (7 == switch_2):
        $ 1332 "Case 7"
        $ 1333 "Sarstedt"
        $ 1334 "'CHANGE THE REFERENCE TO THE FRAME TO MOVE IN'"
        # 'CHANGE THE REFERENCE TO THE FRAME TO MOVE IN'
        $ 1340 "If TASK.ID≟10"
        if (TASK.ID == 10):
          $ 1341 "Frame & Position Params"
          $ 1343 "FRM_Reference = CAM_LM_SSRack"
          FRM_Reference = CAM_LM_SSRack
          $ 1348 "PSE_T≔uLM_SS_PickPlc"
          global PSE_T=uLM_SS_PickPlc
          $ 1349 "PSE_A≔pose_trans(PSE_T, p[0,0,0.1,0,0,0])"
          global PSE_A= pose_trans (PSE_T, p[0,0,0.1,0,0,0])
          $ 1350 "PSE_R≔pose_add(PSE_T, p[0,0,0.1,0,0,0])"
          global PSE_R= pose_add (PSE_T, p[0,0,0.1,0,0,0])
        else:
          $ 1351 "ElseIf TASK.ID≟11"
          if (TASK.ID == 11):
            $ 1352 "FRM_Reference = ULM_SS_Jig"
            FRM_Reference = ULM_SS_Jig
            $ 1353 "PSE_T≔pose_RPY2RotVec(p[0,0,0,0,0,0])"
            global PSE_T=pose_RPY2RotVec(p[0,0,0,0,0,0])
            $ 1354 "PSE_T≔pose_trans(PSE_T, GRP_Offset)"
            global PSE_T=pose_trans(PSE_T, GRP_Offset)
            $ 1355 "PSE_A≔pose_trans(PSE_T, p[0,0,0.1,0,0,0])"
            global PSE_A= pose_trans (PSE_T, p[0,0,0.1,0,0,0])
            $ 1356 "PSE_R≔pose_add(PSE_T, p[0,0,0.2,0,0,0])"
            global PSE_R= pose_add (PSE_T, p[0,0,0.2,0,0,0])
          end
        end
      elif (8 == switch_2):
        $ 1357 "Case 8"
        $ 1358 "NoK"
        $ 1359 "define poses"
        $ 1360 "'NoK'"
        # 'NoK'
        $ 1361 "FRM_Reference=ULM_NoK"
        FRM_Reference=ULM_NoK
        $ 1362 "PSE_T≔pose_RPY2RotVec(p[0,0,0,0,0,0])"
        global PSE_T=pose_RPY2RotVec(p[0,0,0,0,0,0])
        $ 1363 "PSE_A≔pose_trans(PSE_T, p[0,0,0.1,0,0,0])"
        global PSE_A= pose_trans (PSE_T, p[0,0,0.1,0,0,0])
        $ 1364 "PSE_R≔pose_add(PSE_T, p[0,0,0.100,0,0,0])"
        global PSE_R= pose_add (PSE_T, p[0,0,0.100,0,0,0])
      end
    elif (2 == switch_1):
      $ 1365 "Case 2"
      $ 1366 "Centrifuge"
      $ 1367 "'CHANGE THE REFERENCE TO THE FRAME TO MOVE IN'"
      # 'CHANGE THE REFERENCE TO THE FRAME TO MOVE IN'
      $ 1368 "define poses"
      $ 1369 "FRM_Reference≔FRM_Centrifuge"
      global FRM_Reference=FRM_Centrifuge
      $ 1370 "PSE_T≔GRP_Offset"
      global PSE_T=GRP_Offset
      $ 1371 "If Action≟8"
      if (Action == 8):
        $ 1372 "PSE_R≔pose_add(PSE_T, p[0,0,0.250,0,0,0])"
        global PSE_R= pose_add (PSE_T, p[0,0,0.250,0,0,0])
        $ 1373 "PSE_A≔pose_add(PSE_T, p[0,0,0.150,0,0,0])"
        global PSE_A= pose_add (PSE_T, p[0,0,0.150,0,0,0])
      else:
        $ 1374 "ElseIf Action≟7"
        if (Action == 7):
          $ 1375 "PSE_R≔pose_add(PSE_T, p[0,0,0.150,0,0,0])"
          global PSE_R= pose_add (PSE_T, p[0,0,0.150,0,0,0])
          $ 1376 "PSE_A≔pose_add(PSE_T, p[0,0,0.250,0,0,0])"
          global PSE_A= pose_add (PSE_T, p[0,0,0.250,0,0,0])
        end
      end
    elif (3 == switch_1):
      $ 1377 "Case 3"
      $ 1378 "Output"
      $ 1379 "'CHANGE THE REFERENCE TO THE FRAME TO MOVE IN'"
      # 'CHANGE THE REFERENCE TO THE FRAME TO MOVE IN'
      $ 1380 "define poses"
      $ 1381 "FRM_Reference≔Base_const"
      global FRM_Reference=p[0.0,0.0,0.0,0.0,0.0,0.0]
      $ 1382 "PSE_T≔p[0,0,0,0,0,0]"
      global PSE_T=p[0,0,0,0,0,0]
      $ 1383 "PSE_A≔pose_add(PSE_T, p[0,0,0.150,0,0,0])"
      global PSE_A= pose_add (PSE_T, p[0,0,0.150,0,0,0])
      $ 1384 "PSE_R≔pose_add(PSE_T, p[0,0,0.100,0,0,0])"
      global PSE_R= pose_add (PSE_T, p[0,0,0.100,0,0,0])
    elif (5 == switch_1):
      $ 1385 "Case 5"
      $ 1386 "Sarstedt Pickup Table"
      $ 1387 "'CHANGE THE REFERENCE TO THE FRAME TO MOVE IN'"
      # 'CHANGE THE REFERENCE TO THE FRAME TO MOVE IN'
      $ 1388 "Switch JIG"
      switch_2 = JIG
      $ 1389 "Case 7"
      if (7 == switch_2):
        $ 1402 "Sarstedt"
        $ 1403 "'CHANGE THE REFERENCE TO THE FRAME TO MOVE IN'"
        # 'CHANGE THE REFERENCE TO THE FRAME TO MOVE IN'
        $ 1409 "If TASK.ID≟10"
        if (TASK.ID == 10):
          $ 1410 "Frame & Position Params"
          $ 1412 "FRM_Reference = CAM_LM_SSRack"
          FRM_Reference = CAM_LM_SSRack
          $ 1417 "PSE_T≔uLM_SS_PickPlc"
          global PSE_T=uLM_SS_PickPlc
          $ 1418 "PSE_A≔pose_trans(PSE_T, p[0,0,0.1,0,0,0])"
          global PSE_A= pose_trans (PSE_T, p[0,0,0.1,0,0,0])
          $ 1419 "PSE_R≔pose_add(PSE_T, p[0,0,0.1,0,0,0])"
          global PSE_R= pose_add (PSE_T, p[0,0,0.1,0,0,0])
        end
      end
    end
    $ 1426 "Additional check"
    $ 1427 "If  not is_reachable(FRM_Reference,[PSE_A,PSE_A_H,PSE_T,PSE_T_H,PSE_R,PSE_R_H])"
    if (  not  is_reachable(FRM_Reference,[PSE_A,PSE_A_H,PSE_T,PSE_T_H,PSE_R,PSE_R_H])):
      $ 1428 "Error"
      $ 1429 "set_error(ERROR_POSE_NOT_REACHABLE)"
      set_error(ERROR_POSE_NOT_REACHABLE)
      $ 1430 "Action≔0"
      global Action=0
    end
    $ 1431 "'=========='"
    # '=========='
    $ 1432 "Switch Action"
    switch_1 = Action
    $ 1433 "Case 1"
    if (1 == switch_1):
      $ 1434 "Pick"
      $ 1435 "Action_Info≔'pick object'"
      global Action_Info="pick object"
      $ 1436 "do_transition(pose_trans(FRM_Reference, PSE_T), keep_rxry=OBJ_Picked)"
      do_transition( pose_trans (FRM_Reference, PSE_T), keep_rxry=OBJ_Picked)
      $ 1437 "EOAT"
      $ 1438 "If  not OBJ_Picked"
      if (  not  OBJ_Picked):
        $ 1439 "rq_move_and_wait_mm(GRP_Open_Pos)"
         rq_move_and_wait_mm (GRP_Open_Pos)
      end
      $ 1440 "If PSE_A_H≠PSE_Z"
      if (PSE_A_H != PSE_Z):
        $ 1441 "If JNT_Q≠JNT_Z"
        if (JNT_Q != JNT_Z):
          $ 1442 "movej(get_inverse_kin(pose_trans(FRM_Reference, PSE_A_H), qnear=JNT_Q), r=0.050)"
          movej(get_inverse_kin( pose_trans (FRM_Reference, PSE_A_H), qnear=JNT_Q), r=0.050)
        else:
          $ 1443 "Else" "noBreak"
          $ 1444 "movej(pose_trans(FRM_Reference, PSE_A_H), r=0.050)"
          movej( pose_trans (FRM_Reference, PSE_A_H), r=0.050)
        end
      end
      $ 1445 "If PSE_A≠PSE_Z"
      if (PSE_A != PSE_Z):
        $ 1446 "If JNT_Q≠JNT_Z"
        if (JNT_Q != JNT_Z):
          $ 1447 "movej(get_inverse_kin(pose_trans(FRM_Reference, PSE_A), qnear=JNT_Q), r=0.020)"
          movej(get_inverse_kin( pose_trans (FRM_Reference, PSE_A), qnear=JNT_Q), r=0.020)
        else:
          $ 1448 "Else" "noBreak"
          $ 1449 "movej(pose_trans(FRM_Reference, PSE_A), r=0.020)"
          movej( pose_trans (FRM_Reference, PSE_A), r=0.020)
        end
      end
      $ 1450 "MoveL"
      $ 1451 "If PSE_T_H≠PSE_Z"
      if (PSE_T_H != PSE_Z):
        $ 1452 "PSE_T_H" "breakAfter"
        movel(pose_trans(FRM_Reference, PSE_T_H), a=0.5, v=0.4, r=0.01)
      end
      $ 1453 "PSE_T" "breakAfter"
      movel(pose_trans(FRM_Reference, PSE_T), a=0.08, v=0.12)
      $ 1454 "EOAT"
      $ 1455 "rq_set_force_norm(50)"
       rq_set_force_norm (50)
      $ 1456 "rq_close_and_wait()"
       rq_close_and_wait ()
      $ 1457 "OBJ_Picked≔rq_is_object_detected()"
      global OBJ_Picked= rq_is_object_detected ()
      $ 1458 "If  not OBJ_Picked"
      if (  not  OBJ_Picked):
        $ 1459 "set_error(ERROR_NO_OBJECT_TO_PICK)"
        set_error(ERROR_NO_OBJECT_TO_PICK)
      end
      $ 1460 "EXTT"
      $ 1461 "Switch JIG"
      switch_2 = JIG
      $ 1462 "Case 1"
      if (1 == switch_2):
        $ 1463 "3FG"
        $ 1464 "If OBJ_Picked"
        if (OBJ_Picked):
          $ 1465 "Set GRP_3F_Open=On"
          set_standard_digital_out(5, True)
        end
      end
      $ 1466 "If PSE_R_H≠PSE_Z"
      if (PSE_R_H != PSE_Z):
        $ 1467 "PSE_R" "breakAfter"
        movel(pose_trans(FRM_Reference, PSE_R), a=0.5, v=0.4, r=0.01)
        $ 1468 "PSE_R_H" "breakAfter"
        movel(pose_trans(FRM_Reference, PSE_R_H), a=0.5, v=0.4)
      else:
        $ 1469 "Else" "noBreak"
        $ 1470 "PSE_R" "breakAfter"
        movel(pose_trans(FRM_Reference, PSE_R), a=0.5, v=0.4)
      end
    elif (2 == switch_1):
      $ 1471 "Case 2"
      $ 1472 "Place"
      $ 1473 "Action_Info≔'place object'"
      global Action_Info="place object"
      $ 1474 "do_transition(pose_trans(FRM_Reference, PSE_T), keep_rxry=OBJ_Picked)"
      do_transition( pose_trans (FRM_Reference, PSE_T), keep_rxry=OBJ_Picked)
      $ 1475 "EXTT"
      $ 1476 "Switch JIG"
      switch_2 = JIG
      $ 1477 "Case 1"
      if (1 == switch_2):
        $ 1478 "3FG"
        $ 1479 "If OBJ_Picked"
        if (OBJ_Picked):
          $ 1480 "Set GRP_3F_Open=On"
          set_standard_digital_out(5, True)
        end
      end
      $ 1481 "If PSE_A_H≠PSE_Z"
      if (PSE_A_H != PSE_Z):
        $ 1482 "If JNT_Q≠JNT_Z"
        if (JNT_Q != JNT_Z):
          $ 1483 "movej(get_inverse_kin(pose_trans(FRM_Reference, PSE_A_H), qnear=JNT_Q), r=0.050)"
          movej(get_inverse_kin( pose_trans (FRM_Reference, PSE_A_H), qnear=JNT_Q), r=0.050)
        else:
          $ 1484 "Else" "noBreak"
          $ 1485 "movej(pose_trans(FRM_Reference, PSE_A_H), r=0.050)"
          movej( pose_trans (FRM_Reference, PSE_A_H), r=0.050)
        end
      end
      $ 1486 "If PSE_A≠PSE_Z"
      if (PSE_A != PSE_Z):
        $ 1487 "If JNT_Q≠JNT_Z"
        if (JNT_Q != JNT_Z):
          $ 1488 "movej(get_inverse_kin(pose_trans(FRM_Reference, PSE_A), qnear=JNT_Q), r=0.020)"
          movej(get_inverse_kin( pose_trans (FRM_Reference, PSE_A), qnear=JNT_Q), r=0.020)
        else:
          $ 1489 "Else" "noBreak"
          $ 1490 "movej(pose_trans(FRM_Reference, PSE_A), r=0.020)"
          movej( pose_trans (FRM_Reference, PSE_A), r=0.020)
        end
      end
      $ 1491 "MoveL"
      $ 1492 "If PSE_T_H≠PSE_Z"
      if (PSE_T_H != PSE_Z):
        $ 1493 "PSE_T_H" "breakAfter"
        movel(pose_trans(FRM_Reference, PSE_T_H), a=0.5, v=0.4, r=0.01)
      end
      $ 1494 "PSE_T" "breakAfter"
      global move_thread_flag_1494=0
      thread move_thread_1494():
        enter_critical
        move_thread_flag_1494 = 1
        movel(pose_trans(FRM_Reference, PSE_T), a=0.05, v=0.09)
        move_thread_flag_1494 = 2
        exit_critical
      end
      move_thread_flag_1494 = 0
      move_thread_han_1494 = run move_thread_1494()
      while (True):
        local targetTcpDirection=get_target_tcp_speed()
        local stepsToRetract=tool_contact(direction=targetTcpDirection)
        if (stepsToRetract > 0):
          kill move_thread_han_1494
          stopl(0.5)
          $ 1495 "Until (tool_contact_detection)"
          break
        end
        sleep(1.0E-10)
        if (move_thread_flag_1494 > 1):
          join move_thread_han_1494
          break
        end
        sync()
      end
      $ 1496 "Force"
      sleep(0.02)
      zero_ftsensor()
      force_mode(FRM_Reference, [1, 1, 1, 0, 0, 0], [0.0, 0.0, 0.0, 0.0, 0.0, 0.0], 2, [0.1, 0.1, 0.01, 0.3490658503988659, 0.3490658503988659, 0.3490658503988659])
      $ 1497 "PSE_T" "noBreak"
      movel(pose_trans(FRM_Reference, PSE_T), a=0.04, v=0.07)
      end_force_mode()
      stopl(5.0)
      $ 1498 "EXTT"
      $ 1499 "Switch JIG"
      switch_2 = JIG
      $ 1500 "Case 1"
      if (1 == switch_2):
        $ 1501 "3FG"
        $ 1502 "If OBJ_Picked"
        if (OBJ_Picked):
          $ 1503 "Set GRP_3F_Open=Off"
          set_standard_digital_out(5, False)
          $ 1504 "Wait: 0.2"
          sleep(0.2)
        end
      end
      $ 1505 "EOAT"
      $ 1506 "rq_move_and_wait_mm(GRP_Open_Pos)"
       rq_move_and_wait_mm (GRP_Open_Pos)
      $ 1507 "OBJ_Picked≔rq_is_object_detected()"
      global OBJ_Picked= rq_is_object_detected ()
      $ 1508 "If PSE_R_H≠PSE_Z"
      if (PSE_R_H != PSE_Z):
        $ 1509 "PSE_R" "breakAfter"
        movel(pose_trans(FRM_Reference, PSE_R), a=0.5, v=0.4, r=0.01)
        $ 1510 "PSE_R_H" "breakAfter"
        movel(pose_trans(FRM_Reference, PSE_R_H), a=0.5, v=0.4)
      else:
        $ 1511 "Else" "noBreak"
        $ 1512 "PSE_R" "breakAfter"
        movel(pose_trans(FRM_Reference, PSE_R), a=0.5, v=0.4)
      end
    elif (3 == switch_1):
      $ 1513 "Case 3"
      $ 1514 "Push"
      $ 1515 "Action_Info≔'push'"
      global Action_Info="push"
    elif (4 == switch_1):
      $ 1516 "Case 4"
      $ 1517 "Pull"
      $ 1518 "Action_Info≔'pull'"
      global Action_Info="pull"
    elif (6 == switch_1):
      $ 1521 "Case 6"
      $ 1522 "Drop the cap"
      $ 1523 "If JNT_A≠[0,0,0,0,0,0]"
      if (JNT_A != [0,0,0,0,0,0]):
        $ 1524 "MoveJ"
        $ 1525 "JNT_A" "breakAfter"
        movej(JNT_A, a=1.3962634015954636, v=1.7453292519943295, r=0.02)
      else:
        $ 1526 "Else" "noBreak"
        $ 1527 "MoveJ"
        $ 1528 "PSE_A" "breakAfter"
        movej(pose_trans(FRM_Reference, PSE_A), a=1.3962634015954636, v=1.7453292519943295, r=0.02)
      end
      $ 1529 "MoveL"
      $ 1530 "PSE_T" "breakAfter"
      movel(pose_trans(FRM_Reference, PSE_T), a=0.05, v=0.09)
      $ 1531 "'ADD OPEN GRIPPER'"
      # 'ADD OPEN GRIPPER'
      # begin: URCap Program Node
      #   Source: Robotiq_Grippers, 1.8.4.4844, Robotiq Inc.
      #   Type: Gripper
      $ 1532 "Gripper Move10mm (1)"
      if not(gripper_connected[0]):
        popup("Gripper 1 must be connected to run this program.", "No connection", False, True, True)
      end
      if not(rq_is_gripper_activated("1")):
        popup("Gripper 1 is not activated. Go to Installation tab > Gripper to activate it and run the program again.", "Not activated", False, True, True)
      end
      rq_set_pos_spd_for(201, 0, 28, "1")
      rq_wait_pos_spe_for_request(201, 0, 28, "1")
      rq_go_to("1")
      rq_wait("1")
      # end: URCap Program Node
      $ 1533 "PSE_T_H" "breakAfter"
      movel(pose_trans(FRM_Reference, PSE_T_H), a=0.05, v=0.09)
      # begin: URCap Program Node
      #   Source: Robotiq_Grippers, 1.8.4.4844, Robotiq Inc.
      #   Type: Gripper
      $ 1534 "Gripper Move40mm (1)"
      if not(gripper_connected[0]):
        popup("Gripper 1 must be connected to run this program.", "No connection", False, True, True)
      end
      if not(rq_is_gripper_activated("1")):
        popup("Gripper 1 is not activated. Go to Installation tab > Gripper to activate it and run the program again.", "Not activated", False, True, True)
      end
      rq_set_pos_spd_for(63, 0, 28, "1")
      rq_wait_pos_spe_for_request(63, 0, 28, "1")
      rq_go_to("1")
      rq_wait("1")
      # end: URCap Program Node
      $ 1544 "PSE_R" "breakAfter"
      movel(pose_trans(FRM_Reference, PSE_R), a=0.5, v=0.4)
    elif (7 == switch_1):
      $ 1545 "Case 7"
      $ 1546 "Load"
      $ 1547 "Action_Info≔'load object'"
      global Action_Info="load object"
      $ 1548 "do_transition(pose_trans(FRM_Reference, PSE_T), keep_rxry=OBJ_Picked)"
      do_transition( pose_trans (FRM_Reference, PSE_T), keep_rxry=OBJ_Picked)
      $ 1549 "If PSE_A_H≠PSE_Z"
      if (PSE_A_H != PSE_Z):
        $ 1550 "If JNT_Q≠JNT_Z"
        if (JNT_Q != JNT_Z):
          $ 1551 "movej(get_inverse_kin(pose_trans(FRM_Reference, PSE_A_H), qnear=JNT_Q), r=0.050)"
          movej(get_inverse_kin( pose_trans (FRM_Reference, PSE_A_H), qnear=JNT_Q), r=0.050)
        else:
          $ 1552 "Else" "noBreak"
          $ 1553 "movej(pose_trans(FRM_Reference, PSE_A_H), r=0.050)"
          movej( pose_trans (FRM_Reference, PSE_A_H), r=0.050)
        end
      end
      $ 1554 "If PSE_A≠PSE_Z"
      if (PSE_A != PSE_Z):
        $ 1555 "If JNT_Q≠JNT_Z"
        if (JNT_Q != JNT_Z):
          $ 1556 "movej(get_inverse_kin(pose_trans(FRM_Reference, PSE_A), qnear=JNT_Q), r=0.020)"
          movej(get_inverse_kin( pose_trans (FRM_Reference, PSE_A), qnear=JNT_Q), r=0.020)
        else:
          $ 1557 "Else" "noBreak"
          $ 1558 "movej(pose_trans(FRM_Reference, PSE_A), r=0.020)"
          movej( pose_trans (FRM_Reference, PSE_A), r=0.020)
        end
      end
      $ 1559 "MoveL"
      $ 1560 "If PSE_T_H≠PSE_Z"
      if (PSE_T_H != PSE_Z):
        $ 1561 "PSE_T_H" "breakAfter"
        movel(pose_trans(FRM_Reference, PSE_T_H), a=0.5, v=0.4, r=0.01)
      end
      $ 1562 "PSE_T" "breakAfter"
      global move_thread_flag_1562=0
      thread move_thread_1562():
        enter_critical
        move_thread_flag_1562 = 1
        movel(pose_trans(FRM_Reference, PSE_T), a=0.05, v=0.09)
        move_thread_flag_1562 = 2
        exit_critical
      end
      move_thread_flag_1562 = 0
      move_thread_han_1562 = run move_thread_1562()
      while (True):
        local targetTcpDirection=get_target_tcp_speed()
        local stepsToRetract=tool_contact(direction=targetTcpDirection)
        if (stepsToRetract > 0):
          kill move_thread_han_1562
          stopl(0.5)
          $ 1563 "Until (tool_contact_detection)"
          break
        end
        sleep(1.0E-10)
        if (move_thread_flag_1562 > 1):
          join move_thread_han_1562
          break
        end
        sync()
      end
      $ 1564 "Force"
      sleep(0.02)
      zero_ftsensor()
      force_mode(FRM_Reference, [0, 1, 1, 0, 0, 1], [0.0, 0.0, 0.0, 0.0, 0.0, 0.0], 2, [0.1, 0.05, 0.02, 0.3490658503988659, 0.3490658503988659, 3.141592653589793])
      $ 1565 "PSE_T" "noBreak"
      movel(pose_trans(FRM_Reference, PSE_T), a=0.04, v=0.07)
      end_force_mode()
      stopl(5.0)
      $ 1566 "EOAT"
      $ 1567 "rq_move_and_wait_mm(GRP_Open_Pos)"
       rq_move_and_wait_mm (GRP_Open_Pos)
      $ 1568 "OBJ_Picked≔rq_is_object_detected()"
      global OBJ_Picked= rq_is_object_detected ()
      $ 1569 "If PSE_R_H≠PSE_Z"
      if (PSE_R_H != PSE_Z):
        $ 1570 "PSE_R" "breakAfter"
        movel(pose_trans(FRM_Reference, PSE_R), a=0.5, v=0.4, r=0.01)
        $ 1571 "PSE_R_H" "breakAfter"
        movel(pose_trans(FRM_Reference, PSE_R_H), a=0.5, v=0.4)
      else:
        $ 1572 "Else" "noBreak"
        $ 1573 "PSE_R" "breakAfter"
        movel(pose_trans(FRM_Reference, PSE_R), a=0.5, v=0.4)
      end
    elif (8 == switch_1):
      $ 1574 "Case 8"
      $ 1575 "Unload"
      $ 1576 "Action_Info≔'pick object'"
      global Action_Info="pick object"
      $ 1577 "do_transition(pose_trans(FRM_Reference, PSE_T), keep_rxry=OBJ_Picked)"
      do_transition( pose_trans (FRM_Reference, PSE_T), keep_rxry=OBJ_Picked)
      $ 1578 "EOAT"
      $ 1579 "If  not OBJ_Picked"
      if (  not  OBJ_Picked):
        $ 1580 "rq_move_and_wait_mm(GRP_Open_Pos)"
         rq_move_and_wait_mm (GRP_Open_Pos)
      end
      $ 1581 "If PSE_A_H≠PSE_Z"
      if (PSE_A_H != PSE_Z):
        $ 1582 "If JNT_Q≠JNT_Z"
        if (JNT_Q != JNT_Z):
          $ 1583 "movej(get_inverse_kin(pose_trans(FRM_Reference, PSE_A_H), qnear=JNT_Q), r=0.050)"
          movej(get_inverse_kin( pose_trans (FRM_Reference, PSE_A_H), qnear=JNT_Q), r=0.050)
        else:
          $ 1584 "Else" "noBreak"
          $ 1585 "movej(pose_trans(FRM_Reference, PSE_A_H), r=0.050)"
          movej( pose_trans (FRM_Reference, PSE_A_H), r=0.050)
        end
      end
      $ 1586 "If PSE_A≠PSE_Z"
      if (PSE_A != PSE_Z):
        $ 1587 "If JNT_Q≠JNT_Z"
        if (JNT_Q != JNT_Z):
          $ 1588 "movej(get_inverse_kin(pose_trans(FRM_Reference, PSE_A), qnear=JNT_Q), r=0.020)"
          movej(get_inverse_kin( pose_trans (FRM_Reference, PSE_A), qnear=JNT_Q), r=0.020)
        else:
          $ 1589 "Else" "noBreak"
          $ 1590 "movej(pose_trans(FRM_Reference, PSE_A), r=0.020)"
          movej( pose_trans (FRM_Reference, PSE_A), r=0.020)
        end
      end
      $ 1591 "MoveL"
      $ 1592 "If PSE_T_H≠PSE_Z"
      if (PSE_T_H != PSE_Z):
        $ 1593 "PSE_T_H" "breakAfter"
        movel(pose_trans(FRM_Reference, PSE_T_H), a=0.5, v=0.4, r=0.01)
      end
      $ 1594 "PSE_T" "breakAfter"
      movel(pose_trans(FRM_Reference, PSE_T), a=0.08, v=0.12)
      $ 1595 "Force"
      sleep(0.02)
      zero_ftsensor()
      force_mode(FRM_Reference, [1, 1, 0, 0, 0, 0], [0.0, 0.0, 0.0, 0.0, 0.0, 0.0], 2, [0.05, 0.05, 0.1, 0.3490658503988659, 0.3490658503988659, 0.3490658503988659])
      $ 1596 "EOAT" "noBreak"
      $ 1597 "rq_set_force_norm(50)" "noBreak"
       rq_set_force_norm (50)
      $ 1598 "rq_close_and_wait()" "noBreak"
       rq_close_and_wait ()
      $ 1599 "OBJ_Picked≔rq_is_object_detected()" "noBreak"
      global OBJ_Picked= rq_is_object_detected ()
      $ 1600 "If  not OBJ_Picked" "noBreak"
      if (  not  OBJ_Picked):
        $ 1601 "set_error(ERROR_NO_OBJECT_TO_PICK)" "noBreak"
        set_error(ERROR_NO_OBJECT_TO_PICK)
      end
      $ 1602 "If PSE_R_H≠PSE_Z" "noBreak"
      if (PSE_R_H != PSE_Z):
        $ 1603 "PSE_R" "noBreak"
        movel(pose_trans(FRM_Reference, PSE_R), a=0.5, v=0.4, r=0.01)
        $ 1604 "PSE_R_H" "noBreak"
        movel(pose_trans(FRM_Reference, PSE_R_H), a=0.5, v=0.4)
      else:
        $ 1605 "Else" "noBreak"
        $ 1606 "PSE_R" "noBreak"
        movel(pose_trans(FRM_Reference, PSE_R), a=0.5, v=0.4)
      end
      end_force_mode()
      stopl(5.0)
    elif (11 == switch_1):
      $ 1607 "Case 11"
      $ 1608 "Place"
      $ 1609 "Action_Info≔'place object without gripper opening'"
      global Action_Info="place object without gripper opening"
      $ 1610 "do_transition(pose_trans(FRM_Reference, PSE_T), keep_rxry=OBJ_Picked)"
      do_transition( pose_trans (FRM_Reference, PSE_T), keep_rxry=OBJ_Picked)
      $ 1611 "EXTT"
      $ 1612 "Switch JIG"
      switch_2 = JIG
      $ 1613 "Case 1"
      if (1 == switch_2):
        $ 1614 "3FG"
        $ 1615 "If OBJ_Picked"
        if (OBJ_Picked):
          $ 1616 "Set GRP_3F_Open=On"
          set_standard_digital_out(5, True)
        end
      end
      $ 1617 "If PSE_A_H≠PSE_Z"
      if (PSE_A_H != PSE_Z):
        $ 1618 "If JNT_Q≠JNT_Z"
        if (JNT_Q != JNT_Z):
          $ 1619 "movej(get_inverse_kin(pose_trans(FRM_Reference, PSE_A_H), qnear=JNT_Q), r=0.050)"
          movej(get_inverse_kin( pose_trans (FRM_Reference, PSE_A_H), qnear=JNT_Q), r=0.050)
        else:
          $ 1620 "Else" "noBreak"
          $ 1621 "movej(pose_trans(FRM_Reference, PSE_A_H), r=0.050)"
          movej( pose_trans (FRM_Reference, PSE_A_H), r=0.050)
        end
      end
      $ 1622 "If PSE_A≠PSE_Z"
      if (PSE_A != PSE_Z):
        $ 1623 "If JNT_Q≠JNT_Z"
        if (JNT_Q != JNT_Z):
          $ 1624 "movej(get_inverse_kin(pose_trans(FRM_Reference, PSE_A), qnear=JNT_Q), r=0.020)"
          movej(get_inverse_kin( pose_trans (FRM_Reference, PSE_A), qnear=JNT_Q), r=0.020)
        else:
          $ 1625 "Else" "noBreak"
          $ 1626 "movej(pose_trans(FRM_Reference, PSE_A), r=0.020)"
          movej( pose_trans (FRM_Reference, PSE_A), r=0.020)
        end
      end
      $ 1627 "MoveL"
      $ 1628 "If PSE_T_H≠PSE_Z"
      if (PSE_T_H != PSE_Z):
        $ 1629 "PSE_T_H" "breakAfter"
        movel(pose_trans(FRM_Reference, PSE_T_H), a=0.5, v=0.4, r=0.01)
      end
      $ 1630 "PSE_T" "breakAfter"
      global move_thread_flag_1630=0
      thread move_thread_1630():
        enter_critical
        move_thread_flag_1630 = 1
        movel(pose_trans(FRM_Reference, PSE_T), a=0.05, v=0.09)
        move_thread_flag_1630 = 2
        exit_critical
      end
      move_thread_flag_1630 = 0
      move_thread_han_1630 = run move_thread_1630()
      while (True):
        local targetTcpDirection=get_target_tcp_speed()
        local stepsToRetract=tool_contact(direction=targetTcpDirection)
        if (stepsToRetract > 0):
          kill move_thread_han_1630
          stopl(0.5)
          $ 1631 "Until (tool_contact_detection)"
          break
        end
        sleep(1.0E-10)
        if (move_thread_flag_1630 > 1):
          join move_thread_han_1630
          break
        end
        sync()
      end
      $ 1632 "Force"
      sleep(0.02)
      zero_ftsensor()
      force_mode(FRM_Reference, [1, 1, 1, 0, 0, 0], [0.0, 0.0, 0.0, 0.0, 0.0, 0.0], 2, [0.1, 0.1, 0.01, 0.3490658503988659, 0.3490658503988659, 0.3490658503988659])
      $ 1633 "PSE_T" "noBreak"
      movel(pose_trans(FRM_Reference, PSE_T), a=0.04, v=0.07)
      end_force_mode()
      stopl(5.0)
      $ 1634 "EXTT"
      $ 1635 "Switch JIG"
      switch_2 = JIG
      $ 1636 "Case 1"
      if (1 == switch_2):
        $ 1637 "3FG"
        $ 1638 "If OBJ_Picked"
        if (OBJ_Picked):
          $ 1639 "Set GRP_3F_Open=Off"
          set_standard_digital_out(5, False)
          $ 1640 "Wait: 0.2"
          sleep(0.2)
        end
      end
      $ 1641 "EOAT"
      $ 1642 "Comment"
      # Comment
    elif (12 == switch_1):
      $ 1643 "Case 12"
      $ 1644 "Decap"
      $ 1645 "Action_Info≔'decapping'"
      global Action_Info="decapping"
      $ 1646 "Set GRP_3F_Enable=On"
      set_standard_digital_out(4, True)
      $ 1647 "Set GRP_3F_Decap=On"
      set_standard_digital_out(3, True)
      $ 1648 "Force"
      sleep(0.02)
      zero_ftsensor()
      force_mode(tool_pose(), [0, 0, 1, 0, 0, 0], [0.0, 0.0, 5.0, 0.0, 0.0, 0.0], 2, [0.1, 0.1, 0.15, 0.3490658503988659, 0.3490658503988659, 0.3490658503988659])
      $ 1649 "check_decapping(offset=0.015, timeout=5, abort=CMD_Hold)" "noBreak"
      check_decapping(offset=0.015, timeout=5, abort=CMD_Hold)
      end_force_mode()
      stopl(5.0)
      $ 1650 "Set GRP_3F_Decap=Off"
      set_standard_digital_out(3, False)
      $ 1651 "Set GRP_3F_Enable=Off"
      set_standard_digital_out(4, False)
      $ 1652 "MoveL"
      $ 1653 "PSE_R" "breakAfter"
      movel(pose_trans(FRM_Reference, PSE_R), a=0.8, v=0.15)
    elif (13 == switch_1):
      $ 1654 "Case 13"
      $ 1655 "TMR_Barcode: Reset"
      TMR_Barcode = 0
      $ 1656 "Read"
      $ 1657 "TMR_Barcode: Start"
      TMR_Barcode_is_counting = True
      $ 1658 "If TMR_Barcode<PRM_TO_Read_BC"
      global thread_flag_1658=0
      thread Thread_if_1658():
        $ 1659 "KeyenceTrigger"
        $ 1660 "Set OClearResult=HI:Pulse 0.2"
        thread SinglePulse22():
          write_output_boolean_register(2, True)
          sleep(0.2)
          write_output_boolean_register(2, False)
        end
        singlePulse22 = run SinglePulse22()
        $ 1661 "Wait: 0.5"
        sleep(0.5)
        $ 1662 "Set OTriggerBarcode=Off"
        write_output_boolean_register(1, False)
        $ 1663 "Wait: 0.5"
        sleep(0.5)
        $ 1664 "Set OTriggerBarcode=On"
        write_output_boolean_register(1, True)
        $ 1665 "Wait: 0.5"
        sleep(0.5)
        $ 1666 "Preorient"
        $ 1667 "TMR_Barcode: Reset"
        TMR_Barcode = 0
        $ 1668 "If ICmdExctd"
        if (read_input_boolean_register(12)):
          $ 1669 "Set GRP_3F_Decap=On"
          set_standard_digital_out(3, True)
          $ 1670 "Set GRP_3F_Enable=On"
          set_standard_digital_out(4, True)
          $ 1671 "Loop ICmdExctd"
          while (read_input_boolean_register(12)):
            $ 1672 "KeyenceTrigger"
            $ 1673 "Set OClearResult=HI:Pulse 0.1"
            thread SinglePulse23():
              write_output_boolean_register(2, True)
              sleep(0.1)
              write_output_boolean_register(2, False)
            end
            singlePulse23 = run SinglePulse23()
            $ 1674 "Wait: 0.3"
            sleep(0.3)
            $ 1675 "Set OTriggerBarcode=Off"
            write_output_boolean_register(1, False)
            $ 1676 "Wait: 0.3"
            sleep(0.3)
            $ 1677 "Set OTriggerBarcode=On"
            write_output_boolean_register(1, True)
            $ 1678 "Wait: 0.1"
            sleep(0.1)
          end
        end
        $ 1679 "If  not ICmdExctd"
        if (  not  read_input_boolean_register(12)):
          $ 1680 "Set GRP_3F_Decap=On"
          set_standard_digital_out(3, True)
          $ 1681 "Set GRP_3F_Enable=On"
          set_standard_digital_out(4, True)
          $ 1682 "Wait ICmdExctd=HI"
          while (read_input_boolean_register(12) == False):
            sync()
          end
        end
        $ 1683 "Set GRP_3F_Decap=Off"
        set_standard_digital_out(3, False)
        $ 1684 "Set GRP_3F_Enable=Off"
        set_standard_digital_out(4, False)
        $ 1685 "OBJ_Brc_OK≔ True "
        global OBJ_Brc_OK=  True
        thread_flag_1658 = 1
      end
      if (TMR_Barcode<PRM_TO_Read_BC):
        global thread_handler_1658=run Thread_if_1658()
        while (thread_flag_1658 == 0):
          if not(TMR_Barcode<PRM_TO_Read_BC):
            kill thread_handler_1658
            thread_flag_1658 = 2
          else:
            sync()
          end
        end
      else:
        thread_flag_1658 = 2
      end
      if (thread_flag_1658 == 2):
        $ 1686 "Else" "noBreak"
        $ 1687 "exeption"
        $ 1688 "error"
        $ 1690 "OBJ_Brc_OK≔ False "
        global OBJ_Brc_OK=  False
      end
      $ 1691 "Set GRP_3F_Decap=Off"
      set_standard_digital_out(3, False)
      $ 1692 "Set GRP_3F_Enable=Off"
      set_standard_digital_out(4, False)
      $ 1693 "Set OTriggerBarcode=Off"
      write_output_boolean_register(1, False)
    elif (15 == switch_1):
      $ 1694 "Case 15"
      $ 1695 "Detect"
      $ 1696 "Action_Info≔'detect'"
      global Action_Info="detect"
    end
    $ 1697 "'=========='"
    # '=========='
    $ 1698 "PostSettings"
    $ 1699 "'ADD ADDITIONAL CHECKS'"
    # 'ADD ADDITIONAL CHECKS'
  end
  $ 2 "BeforeStart"
  $ 3 "Scripts"
  $ 4 "Script: 001 SCRIPT Errors and Warnings Deifnes V0.2.script"

  #*****************************************************
  # customer          :   UK Essen
  # project name      :   P1132
  #****************************************************
  # controller        :
  # software          :
  #****************************************************
  # author            :   E.Petrichenko
  # Copyright (c)     :   United Robotics Group Health and Food GmbH
  #                       An der Riede 2
  #                       28816 Stuhr
  #                       Germany
  #****************************************************
  # description       :   centrifuge actions for the application
  # version:      	:   0.1
  # created           :   22.08.2024
  # updated           :
  #****************************************************
  # modifications     :
  #
  # date              :
  # name              :
  # reason            :
  #****************************************************


  #################################### VARIABLES DEFINITIONS ###################################

  ERROR_POSE_NOT_REACHABLE = 1002
  ERROR_ROBOT_ARM_NOT_IN_HOME_POSE = 1006
  ERROR_NO_OBJECT_TO_PICK = 1010
  ERROR_NOT_DOCKED = 2003
  ERROR_NOT_REACHABLE_TARGET = 2007
  ERROR_CHARGING_NOT_STARTED = 2008
  ERROR_AMR_WRONG_MODE = 2009
  ERROR_UNKNOWN_POSE = 2010
  ERROR_NO_LANDMARK = 3002
  ERROR_WRONG_ORDER = 4002
  ERROR_CENTRIFUGE_CONNECTION = 5001
  ERROR_CENTRIFUGE_POWER = 5002
  ERROR_CENTRIFUGE = 5003
  ERROR_CENTRIFUGE_LID = 5004
  ERROR_CANNOT_OPEN_HATCH = 5006
  ERROR_CANNOT_CLOSE_HATCH = 5008
  ERROR_CANNOT_ROTATE = 5010
  ERROR_CANNOT_START = 5011
  ERROR_WRONG_KEY_POSE = 5012
  ERROR_MISSIING_CENTRACK = 5013

  WARNING_POSE_NOT_REACHABLE = 1002
  WARNING_BATTERY_LEVEL = 2002
  WARNING_NOT_REACHABLE_TARGET = 2007


  ERROR = struct(
      FLAG = False,
      ID = 0,
      MSG = "")

  WARNING = struct(
      FLAG = False,
      ID = 0,
      MSG = "")


  #################################### FUNCTIONS ###################################

  def set_error(error_id):
      ERROR.ID = error_id
      if (ERROR.ID == 0):
          ERROR.FLAG = False
          ERROR.MSG = ""
      else:
          ERROR.FLAG = True
          if(ERROR.ID == ERROR_POSE_NOT_REACHABLE):
              ERROR.MSG = "Pose is not reachable"
          elif(ERROR.ID == ERROR_NO_OBJECT_TO_PICK):
              ERROR.MSG = "No object to pick"
          elif(ERROR.ID == ERROR_NO_LANDMARK):
              ERROR.MSG = "No landmark detected"
          elif(ERROR.ID == ERROR_ROBOT_ARM_NOT_IN_HOME_POSE):
              ERROR.MSG = "Robot arm cannot go to home pose"
          elif(ERROR.ID == ERROR_AMR_WRONG_MODE):
              ERROR.MSG = "AMR is in the wrong mode"
          elif(ERROR.ID == ERROR_NOT_DOCKED):
              ERROR.MSG = "Could not dock to the charger"
          elif(ERROR.ID == ERROR_NOT_REACHABLE_TARGET):
              ERROR.MSG = "Could not reach the target"
          elif(ERROR.ID == ERROR_CHARGING_NOT_STARTED):
              ERROR.MSG = "Could not start charging"
          elif(ERROR.ID == ERROR_UNKNOWN_POSE):
              ERROR.MSG = "Unknown navigation target"
          elif(ERROR.ID == ERROR_CANNOT_OPEN_HATCH):
              ERROR.MSG = "Centrifuge Cannot open the hatch"
          elif(ERROR.ID == ERROR_CENTRIFUGE_CONNECTION):
              ERROR.MSG = "Cannot reach centrifuge"
          elif (ERROR.ID == ERROR_CANNOT_CLOSE_HATCH):
              ERROR.MSG = "Centrifuge Cannot close the hatch"
          elif (ERROR.ID == ERROR_CANNOT_START):
              ERROR.MSG = "Centrifuge Cannot start"
          elif (ERROR.ID == ERROR_CANNOT_ROTATE):
              ERROR.MSG = "Centrifuge Cannot rotate the rotor"
          elif (ERROR.ID == ERROR_WRONG_ORDER):
              ERROR.MSG = "Wrong parameter was recieved"
          elif (ERROR.ID == ERROR_CENTRIFUGE):
              ERROR.MSG = "Centrifuge is in Error"
          elif (ERROR.ID == ERROR_WRONG_KEY_POSE):
              ERROR.MSG = "Key is in the wrong position"
          elif(ERROR.ID == ERROR_MISSIING_CENTRACK):
              ERROR.MSG = "Missing rack for centrifuge set"
          elif(ERROR.ID == ERROR_CENTRIFUGE_POWER):
              ERROR.MSG = "Centrifuge is turned off"
          elif(ERROR.ID == ERROR_CENTRIFUGE_LID):
              ERROR.MSG = "Lid of the centrifuge is opened"
          else:
              ERROR.MSG = "Unknown code"
          end
          textmsg("ERROR:",ERROR)
      end
  end

  def set_warning(warning_id):
      WARNING.ID = warning_id
      if (WARNING.ID == 0):
          WARNING.FLAG = False
          WARNING.MSG = ""
      else:
          WARNING.FLAG = True
          if(WARNING.ID == WARNING_POSE_NOT_REACHABLE):
              WARNING.MSG = "Pose is not reachable"
          elif(WARNING.ID == WARNING_BATTERY_LEVEL):
              WARNING.MSG = "Batery level dropped to a certain level"
          elif(WARNING.ID == WARNING_NOT_REACHABLE_TARGET):
              WARNING.MSG = "Not reachable location of AMR"
          else:
              WARNING.MSG = "Unknown code"
          end
          textmsg("WARNING:",WARNING)
      end
  end


  def reset_error():
    ERROR.ID = 0
    ERROR.FLAG = False
    ERROR.MSG = ""
  end


  def reset_warning():
      WARNING.ID = 0
      WARNING.FLAG = False
      WARNING.MSG = ""
    end
  $ 5 "Script: SCRIPT uGO V7.11.1.script"
  #*****************************************************
  # customer          :
  # project name      :   Standard Application
  #****************************************************
  # controller        :
  # software          :
  #****************************************************
  # author            :   P. Koehnke
  # Copyright (c)     :   United Robotics Group
  #                       An der Riede 2
  #                       28816 Stuhr
  #                       Germany
  #****************************************************
  # description       :   interface for uGo
  # version:      	:   6.0
  # created           :   21.04.2022
  # updated           :
  #****************************************************
  # modifications     :   add new rpc-functions to interchange more data
  #
  # date              :   2024-02-29
  # name              :   P. Koehnke
  # reason            :   implemtentation of PackML behavoiur in uGO
  #****************************************************
  #****************************************************
  # modifications     :   add reflecting the UID of the uGO task back to uGO
  #
  # date              :   2024-07-02
  # name              :   P. Koehnke
  # reason            :   be sure to finish the right tasks
  #****************************************************

  # available rpc-functions:
  #.on('con_check', (err, _params, callback) => callback(err, this.con_check()))
  #.on('read_input', (err, params, callback) => callback(err, this.read_input(params[0], params[1])))
  #.on('write_output', (err, params, callback) => callback(err, this.write_output(params[0], params[1], params[2])))
  #.on('read_status', (err, params, callback) => callback(err, this.read_status(params[0])))
  #.on('write_status', (err, params, callback) => callback(err, this.write_status(params[0], params[1])))
  #.on('send_template', (err, params, callback) => callback(err, this.receive_state(params[0])))
  #.on('receive_event', (err, params, callback) => callback(err, this.send_event()))
  #.on('send_state', (err, params, callback) => callback(err, this.receive_state(params[0])))
  #.on('send_error', (err, params, callback) => callback(err, this.receive_error(params[0])))
  #.on('NotFound', (methodCalled, params) => LOG.warn('Method "', methodCalled, '" does not exist. ', { params }));

  # =======================================================================
  local IDX_CMD_STOP = 0
  local IDX_CMD_RESET = 1
  local IDX_CMD_START = 2
  local IDX_CMD_HOLD = 3
  local IDX_CMD_UNHOLD = 4
  local IDX_CMD_SUSPEND = 5
  local IDX_CMD_UNSUSPEND = 6
  local IDX_CMD_ABORT = 7
  local IDX_CMD_CLEAR = 8
  local IDX_FNC_FREEDRIVE = 9

  # uGo specific declarations
  global UGO_Request_ID = ""
  global UGO_UNIT_Task = ""
  global UGO_Task_ID = 0
  global UGO_Event = ""
  local UGO_Enable_Control = False
  local UGO = rpc_factory("xmlrpc", "http://192.168.12.120:8080")
  local UGO_Ctrl_Cmd = [False, False, False, False, False, False, False, False, False, False]

  local UGO_AMR_Pos = struct(position_identifier=0, x1=0, x2=0, y1=0, y2=0, theta1=0, theta2=0)
  local UGO_EOAT = struct(object_picked=False)

  def ugo_init(enable=True, rpc_address="http://192.168.12.120:8080"):
      # connection with uGo
      if enable:
          UGO = rpc_factory("xmlrpc", rpc_address)
          UGO_Enable_Control = True
      else:
          UGO_Enable_Control = False
      end
  end

  def ugo_event_controller():
      # interpret the given command and map it to the internal commands
      if UGO_Enable_Control:
          UGO_Event = UGO.receive_event()
      end

      UGO_Ctrl_Cmd[IDX_CMD_STOP] = (UGO_Event == "stop")
      UGO_Ctrl_Cmd[IDX_CMD_RESET] = (UGO_Event == "reset")
      UGO_Ctrl_Cmd[IDX_CMD_START] = (UGO_Event == "start")
      UGO_Ctrl_Cmd[IDX_CMD_HOLD] = (UGO_Event == "hold")
      UGO_Ctrl_Cmd[IDX_CMD_UNHOLD] = (UGO_Event == "un_hold")
      UGO_Ctrl_Cmd[IDX_CMD_SUSPEND] = (UGO_Event == "suspend")
      UGO_Ctrl_Cmd[IDX_CMD_UNSUSPEND] = (UGO_Event == "un_suspend")
      UGO_Ctrl_Cmd[IDX_CMD_ABORT] = (UGO_Event == "abort")
      UGO_Ctrl_Cmd[IDX_CMD_CLEAR] = (UGO_Event == "clear")
      UGO_Ctrl_Cmd[IDX_FNC_FREEDRIVE] = (UGO_Event == "freedrive")

      return UGO_Ctrl_Cmd
  end

  def ugo_translate_pml_state():
      # translate the current PML State to a string
      if (STATE == 1):
          return "STOPPING"
      elif (STATE == 2):
          return "STOPPED"
      elif (STATE == 3):
          return "RESETTING"
      elif (STATE == 4):
          return "IDLE"
      elif (STATE == 5):
          return "STARTING"
      elif (STATE == 6):
          return "EXECUTE"
      elif (STATE == 7):
          return "COMPLETING"
      elif (STATE == 8):
          return "COMPLETE"
      elif (STATE == 9):
          return "HOLDING"
      elif (STATE == 10):
          return "HELD"
      elif (STATE == 11):
          return "UNHOLDING"
      elif (STATE == 12):
          return "SUSPENDING"
      elif (STATE == 13):
          return "SUSPENDED"
      elif (STATE == 14):
          return "UNSUSPENDING"
      elif (STATE == 15):
          return "ABORTING"
      elif (STATE == 16):
          return "ABORTED"
      elif (STATE == 17):
          return "CLEARING"
      else:
          return "UNKNOWN"
      end
  end

  def ugo_update_outputs():
      #Update the outputs to uGo via xmplrpc service
      UGO.write_status("ROB_Skill", UGO_UNIT_Task)
      UGO.write_status("ROB_Battery", AMR_Battery)
      UGO.write_status("ROB_Gripper", OBJ_Picked)
      UGO.send_state(ugo_translate_pml_state(), UGO_UNIT_Task)
      UGO.send_error(ERROR.ID)
      #UGO.send_position(AMR_Position)
  end

  def ugo_get_task():
      # get the actual task to work on
      # added: reflecting the UID of the task back to uGO
      UGO_UNIT_Task = UGO.read_status("DSH_Workflow")
      if (UGO_UNIT_Task != ""):
          UGO_Request_ID = str_sub(UGO_UNIT_Task, 0, 39)
          UGO_Task_ID = to_num(str_sub(UGO_UNIT_Task, 40, 2))
          #ugo_tasks()
          return UGO_Task_ID
      else:
          return 0
      end
  end

  def ugo_pml_stopping():
      return True
  end

  def ugo_pml_resetting():
      ugo_get_task()
      if (UGO_UNIT_Task == ""):
          UGO_Request_ID = ""
          UGO_Task_ID = 0
          return True
      end
      return False
  end

  def ugo_pml_starting():
      #UGO_Task_Content = UGO.receive_task()
      return (UGO_UNIT_Task != "")
  end

  def ugo_pml_holding():
      return True
  end

  def ugo_pml_unholding():
      return True
  end

  def ugo_pml_suspending():
      return True
  end

  def ugo_pml_unsuspending():
      return True
  end

  def ugo_pml_completing():
      return True
  end

  def ugo_pml_aborting():
      return True
  end

  def ugo_pml_clearing():
      return True
  end

  # =======================================================================
  # end of uGO script
  # =======================================================================
  $ 7 "Script: SCRIPT PackML V1.2.1.script"
  # PackML

  IO_ADDRESS_CMD_STOP = 1
  IO_ADDRESS_CMD_RESET = 7
  IO_ADDRESS_CMD_START = 0

  EXT_ADDRESS_CMD_STOP = 0
  EXT_ADDRESS_CMD_RESET = 1
  EXT_ADDRESS_CMD_START = 2
  EXT_ADDRESS_CMD_HOLD = 3
  EXT_ADDRESS_CMD_UNHOLD = 4
  EXT_ADDRESS_CMD_SUSPEND = 5
  EXT_ADDRESS_CMD_UNSUSPEND = 6
  EXT_ADDRESS_CMD_ABORT = 7
  EXT_ADDRESS_CMD_CLEAR = 8
  EXT_ADDRESS_FNC_FREEDRIVE = 9

  global EXT_CtrlCmd = [False, False, False, False, False, False, False, False, False, False]

  EXT_Control_by = "uGO"

  global CMD_Abort = False
  global CMD_Clear = False
  global CMD_Stop = False
  global CMD_Reset = False
  global CMD_Start = False
  global CMD_Hold = False
  global CMD_Unhold = False
  global CMD_Suspend = False
  global CMD_Unsuspend = False
  global FNC_Freedrive = False

  CND_Suspend = False         # condition for suspend command
  CND_Unsuspend = False       # condition for unsuspend command

  thread Get_Pml_Command():
      while (True):
          if (EXT_Control_by == "uGO"):
              EXT_CtrlCmd = ugo_event_controller()
          elif (EXT_Control_by == "Leitsystem"):
              # EXT_CtrlCmd = Leitsystem
          end
          # ---------- Abort ---------- #
          if ((not STATE == 15) and (not STATE == 16) and EXT_CtrlCmd[EXT_ADDRESS_CMD_ABORT]):
              CMD_Abort = True
              CMD_Stop = False
          elif ((STATE == 17) and not EXT_CtrlCmd[EXT_ADDRESS_CMD_ABORT]):
              CMD_Abort = False
          end
          # ---------- Stop ---------- #
          if ((not STATE == 1) and (not STATE == 2) and (get_standard_digital_in(IO_ADDRESS_CMD_STOP) or EXT_CtrlCmd[EXT_ADDRESS_CMD_STOP])):
              CMD_Stop = True
              if get_standard_digital_in(IO_ADDRESS_CMD_STOP):
                  log_state("Stop command by pushbutton")
              elif EXT_CtrlCmd[EXT_ADDRESS_CMD_STOP]:
                  log_state("Stop command by external control")
              end
          elif (STATE == 2) and (not get_standard_digital_in(IO_ADDRESS_CMD_STOP)) and (not EXT_CtrlCmd[EXT_ADDRESS_CMD_STOP]):
              CMD_Stop = False
          end
          CMD_Hold = (STATE == 6 or STATE == 10) and not CMD_Stop and (ERROR.FLAG or EXT_CtrlCmd[EXT_ADDRESS_CMD_HOLD])
          CMD_Reset = (STATE == 2 or STATE == 8) and not CMD_Stop and (read_input_boolean_register(5) or EXT_CtrlCmd[EXT_ADDRESS_CMD_RESET])
          CMD_Start = (STATE == 4) and not CMD_Stop and (get_standard_digital_in(IO_ADDRESS_CMD_START) or EXT_CtrlCmd[EXT_ADDRESS_CMD_START])
          CMD_Unhold = (STATE == 10) and not CMD_Stop and (get_standard_digital_in(IO_ADDRESS_CMD_START) or EXT_CtrlCmd[EXT_ADDRESS_CMD_UNHOLD])
          CMD_Suspend = (STATE == 6) and not CMD_Stop and (CND_Suspend or EXT_CtrlCmd[EXT_ADDRESS_CMD_SUSPEND])
          CMD_Unsuspend = (STATE == 13) and not CMD_Stop and (CND_Unsuspend or EXT_CtrlCmd[EXT_ADDRESS_CMD_UNSUSPEND])
          CMD_Clear = (STATE == 16) and EXT_CtrlCmd[EXT_ADDRESS_CMD_CLEAR]
          FNC_Freedrive = (STATE == 10) and EXT_CtrlCmd[EXT_ADDRESS_FNC_FREEDRIVE]
          sleep(0.1)
      end
  end

  thread_pml_command_handler = run Get_Pml_Command()

  def command_manager(external_control="uGO", cond_suspend=False, cond_unsuspend=False):

      EXT_Control_by = external_control
      CND_Suspend = cond_suspend
      CND_Unsuspend = cond_unsuspend

      if (CMD_Abort and STATE != 15 and STATE != 16):
          STATE = 15
      elif (CMD_Stop and STATE != 1 and STATE != 2):
          STATE = 1
      end
      return False
  end

  def stopping():
      if (EXT_Control_by == "uGO"):
          return ugo_pml_stopping()
      elif (EXT_Control_by == "Leitsystem"):
          # EXT_CtrlCmd = Leitsystem
      else:
          return True
      end
      return False
  end

  def resetting():
      if (EXT_Control_by == "uGO"):
          return ugo_pml_resetting()
      elif (EXT_Control_by == "Leitsystem"):
          # EXT_CtrlCmd = Leitsystem
      else:
          return True
      end
      return False
  end

  def starting():
      if (EXT_Control_by == "uGO"):
          return ugo_pml_starting()
      elif (EXT_Control_by == "Leitsystem"):
          # EXT_CtrlCmd = Leitsystem
      else:
          return True
      end
      return False
  end

  def holding():
      if (EXT_Control_by == "uGO"):
          return ugo_pml_holding()
      elif (EXT_Control_by == "Leitsystem"):
          # EXT_CtrlCmd = Leitsystem
      else:
          return True
      end
      return False
  end

  def unholding():
      if (EXT_Control_by == "uGO"):
          return ugo_pml_unholding()
      elif (EXT_Control_by == "Leitsystem"):
          # EXT_CtrlCmd = Leitsystem
      else:
          return True
      end
      return False
  end

  def suspending():
      if (EXT_Control_by == "uGO"):
          return ugo_pml_suspending()
      elif (EXT_Control_by == "Leitsystem"):
          # EXT_CtrlCmd = Leitsystem
      else:
          return True
      end
      return False
  end

  def unsuspending():
      if (EXT_Control_by == "uGO"):
          return ugo_pml_unsuspending()
      elif (EXT_Control_by == "Leitsystem"):
          # EXT_CtrlCmd = Leitsystem
      else:
          return True
      end
      return False
  end

  def completing():
      if (EXT_Control_by == "uGO"):
          return ugo_pml_completing()
      elif (EXT_Control_by == "Leitsystem"):
          # EXT_CtrlCmd = Leitsystem
      else:
          return True
      end
      return False
  end

  def aborting():
      if (EXT_Control_by == "uGO"):
          return ugo_pml_aborting()
      elif (EXT_Control_by == "Leitsystem"):
          # EXT_CtrlCmd = Leitsystem
      else:
          return True
      end
      return False
  end

  def clearing():
      if (EXT_Control_by == "uGO"):
          return ugo_pml_clearing()
      elif (EXT_Control_by == "Leitsystem"):
          # EXT_CtrlCmd = Leitsystem
      else:
          return True
      end
      return False
  end
  $ 8 "Script: SCRIPT Utility V5.5.script"
  #*****************************************************
  # customer          :   tbd
  # project name      :   tbd
  #****************************************************
  # controller        :
  # software          :
  #****************************************************
  # author            :   P. Koehnke (+49 1628859904; p.koehnke@unitedrobotics.group)
  # Copyright (c)     :   United Robotics Group Health and Food GmbH
  #                       An der Riede 2
  #                       28816 Stuhr
  #                       Germany
  #****************************************************
  # description       :   utility programs for the application
  # version:      	:   3.1
  # created           :   30.01.2023
  # updated           :
  #****************************************************
  # modifications     :   get_tool_free_pose_2(), get_index_from_list()
  #
  # date              :   05.01.2024
  # name              :   PK
  # reason            :
  #****************************************************

  def found_in_matrix(data, req_id, req_idx):
      local id = -1
      local dimensions = size(data)
      local loop_dataset = 0

      while (id != req_id and loop_dataset < dimensions[0]):
          id = data[loop_dataset, 0]
          if (id == req_id):
              return data[loop_dataset, req_idx]
          else:
              loop_dataset = loop_dataset + 1
          end
      end
  end

  def found_in_list(value, list):
      local idx = 0

      while (idx < length(list)):
          if (value == list[idx]):
              return True
          end
          idx = idx + 1
      end
      return False
  end

  def get_index_from_list(list, value = -1):
      local idx = 0

      while (idx < length(list)):
          if (value == -1):
              if (list[idx] != 0):
                  return idx
              end
          else:
              if (list[idx] == value):
                  return idx
              end
          end
          idx = idx + 1
      end
      return -1
  end

  def find_object_by_type(list, type=0):
      local object = list[0]
      local i = 0

      while i < length(list):
          object = list[i]
          if object.type == type:
              return object
          end
          i = i + 1
      end
  end

  def pose_RPY2RotVec(pose):
      local rotvec = rpy2rotvec([d2r(pose[3]), d2r(pose[4]), d2r(pose[5])])
      return p[pose[0], pose[1], pose[2], rotvec[0], rotvec[1], rotvec[2]]
  end

  def pose_RotVec2RPY(pose):
      local rpy = rotvec2rpy([pose[3], pose[4], pose[5]])
      return p[pose[0], pose[1], pose[2], r2d(rpy[0]), r2d(rpy[1]), r2d(rpy[2])]
  end

  def swivel(frame_ref, angles = [0, 0, 0], pose = p[0, 0, 0, 0, 0, 0]):

      local rpy_ref = [0, 0, 0]
      local rpy_new = [0, 0, 0]
      local rotvec_new = [0, 0, 0]
      local pose_from = p[0, 0, 0, 0, 0, 0]
      local pose_to = p[0, 0, 0, 0, 0, 0]
      local i = 0

      if (pose == p[0, 0, 0, 0, 0, 0]):
          pose_to = pose_trans(pose_inv(frame_ref), get_actual_tcp_pose())
      else:
          pose_to = pose
      end

      rpy_ref = rotvec2rpy(frame_ref[3], frame_ref[4], frame_ref[5])

      while (i < 3):
          rpy_new[i] = rpy_ref[i] + d2r(angles[i])
          i = i + 1
      end

      rotvec_new = rpy2rotvec(rpy_new)
      pose_from = p[0, 0, 0, rotvec_new[0], rotvec_new[1], rotvec_new[2]]
      pose_to = p[pose_to[0], pose_to[1], pose_to[2], rotvec_new[0], rotvec_new[1], rotvec_new[2]]

      return pose_trans(pose_from, pose_to)
  end

  def get_random_pose(pose_ref, mode = "", range_max = [0, 0, 0]):
      # modi: "cubic", "rotation"
      # getting a random pose in the x/y-plane. range can be set for each
      # translation and rotation.
      local rpy_random = [0, 0, 0]
      local rotvec_random = [0, 0, 0]
      local pose_random = pose_ref
      local i = 0

      if (mode == "cubic"):
          # cubic mode: random pose takes only x, y and z
          i = 0
          while (i < 3):
              pose_random[i] = pose_ref[i] + range_max[i] * (random() - 0.5)
              i = i + 1
          end
          return pose_random

      elif (mode == "rotation"):
          i = 0
          while (i < 3):
              rpy_random[i] = d2r(range_max[i]) * (random() - 0.5)
              i = i + 1
          end
          rotvec_random = rpy2rotvec(rpy_random)
          pose_random = pose_trans(p[0, 0, 0, rotvec_random[0], rotvec_random[1], rotvec_random[2]], pose_ref)
          return pose_random

      else:
          # unknown mode, return pose_ref
          return pose_ref
      end
  end

  def get_pattern_pos_rectangle(counter, direction, pattern, patterninc = [0, 0], patternsize = [0, 0]):
      # defines the position inside a rectangular pattern
      # pattern describes, how many objects are in x-direction and how many in y-direction [x, y]
      # patternsize will give the total length of each direction [x, y]
      local X_Fac = 0
      local Y_Fac = 0
      local max = pattern[0] * pattern[1]
      local i = 0

      if (1 > counter or counter > max):
          counter = 1
      end

      if pattern[0] == 0:
          pattern[0] = 1
      end

      if pattern[1] == 0:
          pattern[1] = 1
      end

      if (direction == "Y" or direction == "y"):
          X_Fac = floor((counter - 1) / pattern[1])
          Y_Fac = (counter - 1) % pattern[1]
      elif (direction == "X" or direction == "x"):
          X_Fac = (counter - 1) % pattern[0]
          Y_Fac = floor((counter - 1) / pattern[0])
      end

      if patternsize != [0, 0]:
          while i < 2:
              if pattern[i] > 1:
                  patterninc[i] = patternsize[i] / (pattern[i] - 1)
              end
              i = i + 1
          end
      end

      return p[X_Fac * patterninc[0], Y_Fac * patterninc[1], 0, 0, 0, 0]
  end

  def get_pattern_pos_circle(counter, radius, angle, direction, pattern, patternsize = [0, 0]):
      # get the patternpos for a circular pattern through a counter
      # need the radius and the angle in radiants
      local X_Fac = 0
      local Y_Fac = 0
      local rad_bow = 0
      local radius_cal = 0
      local ref = p[0, 0, 0, 0, 0, 0]

      if pattern[0] == 0:
          pattern[0] = 1
      end

      if pattern[1] == 0:
          pattern[1] = 1
      end

      if (direction == "Y" or direction == "y"):
          X_Fac = floor((counter - 1) / pattern[1])
          Y_Fac = (counter - 1) % pattern[1]
      elif (direction == "X" or direction == "x"):
          X_Fac = (counter - 1) % pattern[0]
          Y_Fac = floor((counter - 1) / pattern[0])
      end

      # the opening angle will be calculated in x-direction
      # works only between -90 and 90 degree
      if pattern[0] > 1:
          rad_bow = - angle / (pattern[0] - 1) * X_Fac + angle / 2
      end

      if (counter % 2 == 0 and pattern[1] > 1):
          radius_cal = radius - patternsize[1] / (pattern[1])
      else:
          radius_cal = radius + patternsize[1] / (pattern[1])
      end
      ref = p[0, radius_cal, 0, 0, 0, 0]

      return p[ref[0] * cos(rad_bow) - ref[1] * sin(rad_bow), (ref[0] * sin(rad_bow) + ref[1] * cos(rad_bow)) - radius, 0, 0, 0, 0]
  end

  def get_pattern_counter(pose, direction, pattern, patterninc = [0, 0], patternsize = [0, 0]):
      # returns the counter for a pattern from a given cartesian pose
      local patternpose = p[pose[0], pose[1], 0, 0, 0, 0]
      local X_Fac = 0
      local Y_Fac = 0
      local i = 0

      if patternsize != [0, 0]:
          while i < 2:
              if pattern[i] > 1:
                  patterninc[i] = patternsize[i] / (pattern[i] - 1)
              else:
                  pattern[i] = 0
              end
              i = i + 1
          end
      end

      # calculation of the counter in the desired axis-direction
      if (direction == "x" or direction == "X"):
          if patterninc[0] > 0:
              X_Fac = ceil((patternpose[0] + patterninc[0] / 2) / patterninc[0])
              if X_Fac < 0:
                  X_Fac = 0
              end
          end
          if patterninc[1] > 0:
              Y_Fac = floor((patternpose[1] + patterninc[1] / 2) / patterninc[1])
              if Y_Fac < 0:
                  Y_Fac = 0
            end
          end
          return Y_Fac * pattern[0] + X_Fac
      elif (direction == "y" or direction == "Y"):
          if patterninc[0] > 0:
              X_Fac = floor((patternpose[0] + patterninc[0] / 2) / patterninc[0])
          end
          if patterninc[1] > 0:
              Y_Fac = ceil((patternpose[1] + patterninc[1] / 2) / patterninc[1])
          end
          return X_Fac * pattern[1] + Y_Fac
      end
  end

  def get_plc_reg(mod_sig_name):
      return integer_to_binary_list(modbus_get_signal_status(mod_sig_name))
  end

  def set_plc_reg(mod_sig_name, mod_sig_list):
      modbus_set_output_register(mod_sig_name, binary_list_to_integer(mod_sig_list), False)
  end

  def check_decapping(offset = 0, timeout = 5, abort = False):
      # checken, ob der Deckel schon ab ist
      local start = get_actual_tcp_pose()
      local current_offset = 0
      local timecounter = 0
      while (current_offset < offset and not abort):
          current_offset = pose_dist(start, get_actual_tcp_pose())
          timecounter = timecounter + 1
          if (timecounter * 0.5 == timeout):
              break
          end
          sleep(0.5)
      end
      stopl(0.5)
  end

  def check_capping(torque = 0):
      # checken, wann der Deckel verschraubt ist
      force_mode(get_actual_tcp_pose(), [0, 0, 1, 0, 0, 0], [0, 0, -2.0, 0, 0, 0], 2, [0, 0, 0.100, 0, 0, 0])
  end

  def is_reachable(frame, poses, offsets = [0, 0, 0]):
      local idx = 0
      local pose = p[0, 0, 0, 0, 0, 0]

      while (idx < length(poses)):
          pose = poses[idx]
          pose[0] = pose[0] + offsets[0]
          pose[1] = pose[1] + offsets[1]
          pose[2] = pose[2] + offsets[2]

          if pose != p[0, 0, 0, 0, 0, 0]:
              if (not get_inverse_kin_has_solution(pose_trans(frame, pose))):
                  textmsg(str_cat(str_cat("Pose ", to_str(idx + 1)), " is not reachable"))
                  return False
              end
          end
          idx = idx + 1
      end
      return True
  end

  def is_within_limits(frame, poses, offsets = [0, 0, 0]):
      local idx = 0
      local pose = p[0, 0, 0, 0, 0, 0]

      while (idx < length(poses)):
          pose = poses[idx]
          pose[0] = pose[0] + offsets[0]
          pose[1] = pose[1] + offsets[1]
          pose[2] = pose[2] + offsets[2]

          if is_reachable(frame = frame, poses = poses, offsets = offsets):
              if (not is_within_safety_limits(get_inverse_kin(pose_trans(frame, pose), get_actual_joint_positions()))):
                  textmsg(str_cat(str_cat("Pose ", to_str(idx + 1)), "is out of joint limits"))
                  return False
              else:
                  idx = idx + 1
              end
          else:
              return False
          end
      end
      return True
  end


  def string_to_list(string, separator = "," , endDelimiter = ";" , capacity = 50):
      local string_length = str_len(string)
      local list_out = make_list(length = elements_in_string(string), initial_value = -1, capacity = capacity)
      local cnt = 0
      local idx = 0

      while cnt < string_length-1 :
        textmsg("new loop")
        textmsg(to_str(idx))
        local sepAt = str_find(string, separator, cnt)
        textmsg(to_str(sepAt))
        if sepAt < 0 :
            sepAt = str_find(string, endDelimiter, cnt)
        end
        list_out[idx] = to_num(str_sub(string, cnt, sepAt-cnt))
        idx = idx +1
        cnt = sepAt + 1
      end

      return list_out
  end

  def elements_in_string(string, separator = "," , endDelimiter = ";" , capacity = 50):
     local string_length = str_len(string)
      local len = 0
      local sepAt = 0

      while sepAt < string_length-1 and sepAt>=0 :
        local sepAt = str_find(string, separator, sepAt+1)
        len = len +1
      end

      return len
  end
  $ 9 "Script: SCRIPT uML Lights V1.2.script"

  #****************************************************
  # product           : uLabMobile
  # language          : urscript
  #****************************************************
  # author            :   D.Kreugel
  # Copyright (c)     :   United Robotics Group
  #                       An der Riede 2
  #                       28816 Stuhr
  #                       Germany
  #****************************************************
  # description       :   led controls for uLabMobile
  # version:      	:   1.2
  # created           :   09.08.2024
  # updated           :
  #****************************************************
  # modifications     :   changed conditions to switch lights (not only pml state but also charging state)
  #
  # date              :   09.08.2024
  # name              :   PK
  # reason            :   due to the change in project P1117, we run to often through every state. This leads to to much colorchanges
  #****************************************************

  # HARDWARE CONFIGURATION
  LED_GREEN = struct(type="CO",id=5)
  LED_RED = struct(type="CO",id=6)
  LED_BLUE = struct(type="CO",id=7)

  def set_output(type,id,state=True):
      if(type=="CO"):
          set_configurable_digital_out(id,state)
      elif(type=="DO"):
          set_standard_digital_out(id,state)
      end
  end

  def led_red_on():
      set_output(LED_RED.type,LED_RED.id,True)
  end

  def led_red_off():
      set_output(LED_RED.type,LED_RED.id,False)
  end

  def led_green_on():
      set_output(LED_GREEN.type,LED_GREEN.id,True)
  end

  def led_green_off():
      set_output(LED_GREEN.type,LED_GREEN.id,False)
  end

  def led_blue_on():
      set_output(LED_BLUE.type,LED_BLUE.id,True)
  end

  def led_blue_off():
      set_output(LED_BLUE.type,LED_BLUE.id,False)
  end


  # COLOR MIX
  def color_blue():
      led_blue_on()
      led_green_off()
      led_red_off()
  end

  def color_red():
      led_blue_off()
      led_green_off()
      led_red_on()
  end

  def color_green():
      led_blue_off()
      led_green_on()
      led_red_off()
  end

  def color_yellow():
      led_blue_off()
      led_green_on()
      led_red_on()
  end

  def color_lightblue():
      led_blue_on()
      led_green_on()
      led_red_off()
  end

  def color_violet():
      led_blue_on()
      led_green_off()
      led_red_on()
  end

  def color_white():
      led_blue_on()
      led_green_on()
      led_red_on()
  end

  def led_off():
      led_blue_off()
      led_green_off()
      led_red_off()
  end

